(* IEC 61131-3 sources: daoli-st-library/DL_Process (part 56) *)

(* ---- FB_DL_TireCureBlowdownWatch.st ---- *)
(*
  Name: FB_DL_TireCureBlowdownWatch
  Category: DL_Process
  Version: 1.0.0
  Round: R91 / 2026-11-25
  开源溯源：clean-room 自研（族 轮胎硫化，ST 开源生态实测 0 命中，无外部代码引入）
  功能：1) 按固定观察窗累计两个量：冷凝水总量 _fAccumKg 与排凝阀动作次数 _iAccumAct，
           窗口到点后按「单位动作排水量」比对：
           ratio = 累计冷凝水 / (动作次数 × 单次期望排水量)。
        2) 双向故障判别：
           ① 比值过高（> fBlockRatio）或窗口内动作次数为零而冷凝水已超限 → 判排凝阀堵塞（码 0322 / 0324），
              即水积在腔内排不出去，会稀释硫化温度场并造成胶囊局部过冷；
           ② 比值过低（< fLeakRatio）→ 判排凝阀泄漏（码 0323），即阀频繁动作但排水极少，
              说明阀芯未关严、蒸汽直排，属能耗与安全问题。
        3) 窗口自复位由 TON 的 IN := xEnable AND NOT tonWin.Q 驱动（R188），
           窗口到点仅置 Q 一拍，用于「判定 + 清累计」的一次性动作，不靠外部沿清零。
  边界条件：1) 非有限值闸：冷凝水量、期望排水量、两个比值阈值、窗口先过
           NOT(x > -DL_BIG AND x < DL_BIG)，同时拦 NaN 与 Inf；命中即锁码 0326 进故障相，
           绝不把 NaN 累加进窗口（NaN 一旦进入累计器，整个窗口乃至后续窗口永久污染，R19）。
        2) 分母零闸：比值式分母 = 动作次数 × 单次期望排水量，动作次数为零时走独立判据（码 0324），
           单次期望排水量 fExpectKgPerAct 必须 > DL_EPS 否则锁码 0325（判据全体失效）。
        3) 阈值域闸：须满足 0.0 < fLeakRatio < fBlockRatio，否则两向判据重叠、必有一向永不触发，
           越域锁码 0325。
        4) 累计器安全：非有限值命中时把两个累计器一并清零（码 0326 已锁存），
           并中止本窗口的判定，防污染值跨窗口传播。
        5) 定时器周期刷新（R7）：窗口 TON 与两个边沿实例全部在 CASE 之外无条件调用。
        6) 故障解除路径：故障相内 xReset 上升沿 AND NOT xFault AND 入参/组态合法 → 清锁存回正常，
           回正常后窗口与累计器全部重新起算（不自恢复）。
        7) 状态机兜底：CASE 全态覆盖 + ELSE 强制回故障相并置码 0328、清全部输出。
        8) 输出安全初值（R25）：xBlocked / xLeaking 初值 FALSE，fRatioPct 初值 0.0，正常相显式赋值。
  量纲自证：ratio = (kg) / (无因次 * kg) = 无因次 [-]；fRatioPct = 无因次 * 100 = 百分数 [%]；
           fAccumKg 为累计质量 [kg]，nAccumAct 为动作次数（计数，无量纲）[count]。
  码表 Error codes（本件子带 0091_032x，故障级一律 3 行内置 _uFault/_bFault/_eState）:
    16#0091_0321 信息级：观察窗累计中，尚未判定（不置故障位）
    16#0091_0322 故障级：排凝阀堵塞（单位动作排水量比值过高）
    16#0091_0323 故障级：排凝阀泄漏（单位动作排水量比值过低，蒸汽直排）
    16#0091_0324 故障级：窗口内动作次数为零但冷凝水超限（阀未动作）
    16#0091_0325 故障级：组态越域（期望排水量/比值阈值/窗口非法）
    16#0091_0326 故障级：入参非有限（NaN 或 Inf），累计器已清
    16#0091_0327 故障级：外部故障输入 xFault
    16#0091_0328 故障级：状态机落 ELSE 兜底（非法相位 ID）

  修订历史 Revision :
    2026-11-25  v1.0.0  R91 首版
*)

TYPE E_DL_TcsBlowdownState :
(
    eTcsBdNormal  := 0,     // 正常：窗口比值在带内 / Normal, window ratio within the band
    eTcsBdBlocked := 10,    // 排凝阀堵塞：水排不出去 / Blocked blowdown valve, water cannot be discharged
    eTcsBdLeaking := 20,    // 排凝阀泄漏：蒸汽直排 / Leaking blowdown valve, steam blows through
    eTcsBdFault   := 90     // 故障：入参/组态非法，锁存待解除 / Fault, invalid input, latched
);
END_TYPE

FUNCTION_BLOCK FB_DL_TireCureBlowdownWatch
VAR_INPUT
    xEnable         : BOOL;   // 监视使能 [bool] / Monitoring enable [bool]
    xReset          : BOOL;   // 故障复位（上升沿有效）[bool] / Fault reset, rising edge [bool]
    xFault          : BOOL;   // 外部故障汇总 [bool] / External fault aggregate [bool]
    xCyclePulse     : BOOL;   // 周期完成脉冲（每个模压周期一个脉冲）[bool] / Cycle-complete pulse [bool]
    fCondensateKg   : REAL;   // 本周期冷凝水量增量 [kg] / Condensate increment of this cycle [kg]
    nActCount       : INT;    // 本周期排凝阀动作次数 [count] / Blowdown valve actuations this cycle [count]
    fExpectKgPerAct : REAL;   // 单次动作期望排水量 [kg/act] / Expected discharge per actuation [kg/act]
    fBlockRatio     : REAL;   // 堵塞判定比值上限 [-] / Blockage upper ratio limit [-]
    fLeakRatio      : REAL;   // 泄漏判定比值下限 [-] / Leakage lower ratio limit [-]
    tWindow         : TIME;   // 观察窗时长 [TIME] / Observation window duration [TIME]
END_VAR
VAR_OUTPUT
    fRatioPct       : REAL;   // 窗口单位动作排水量比值（百分数显示）[%] / Window ratio, percent display [%]
    fAccumKg        : REAL;   // 窗口累计冷凝水量 [kg] / Accumulated condensate in the window [kg]
    nAccumAct       : INT;    // 窗口累计动作次数 [count] / Accumulated actuations in the window [count]
    xBlocked        : BOOL;   // 堵塞标志 [bool] / Blockage flag [bool]
    xLeaking        : BOOL;   // 泄漏标志 [bool] / Leakage flag [bool]
    xWindowDone     : BOOL;   // 窗口到点脉冲（单拍）[bool] / Window-complete single-shot flag [bool]
    eState          : E_DL_TcsBlowdownState;   // 状态出口，段尾单点映射 / State outlet, single-point mapped
    nErrId          : UDINT;  // 事件码，0 = 无事件 / Event code, 0 = none
END_VAR
VAR
    tonWin          : TON;    // 观察窗定时（自复位由 IN 取反驱动，R188）[TIME] / Observation window timer
    rtCycle         : R_TRIG; // 周期脉冲上升沿检测 [bool] / Cycle pulse rising edge detector
    rtReset         : R_TRIG; // 复位上升沿检测 [bool] / Reset rising edge detector
    _eState         : E_DL_TcsBlowdownState := E_DL_TcsBlowdownState.eTcsBdNormal;   // 内部相位（CASE 唯一写入目标）
    _fAccumKg       : REAL := 0.0;   // 窗口累计冷凝水量 [kg] / Accumulated condensate [kg]
    _iAccumAct      : INT := 0;      // 窗口累计动作次数 [count] / Accumulated actuations [count]
    _fRatioRaw      : REAL := 0.0;   // 窗口比值原始值（无因次）[-] / Raw window ratio [-]
    _fRatioRawPct   : REAL := 0.0;   // 窗口比值百分数原始值 [%] / Raw window ratio in percent [%]
    _bFinOk         : BOOL := FALSE; // 实值入参有限性总闸结果 / Finiteness gate aggregate result
    _bCfgOk         : BOOL := FALSE; // 阈值与窗口组态域闸结果 / Threshold and window domain gate result
    _bJudgeThis     : BOOL := FALSE; // 本拍需执行窗口判定（窗口到点）[bool] / Judge this cycle flag
    _bBlockedL      : BOOL := FALSE; // 堵塞锁存位 [bool] / Latched blockage flag
    _bLeakingL      : BOOL := FALSE; // 泄漏锁存位 [bool] / Latched leakage flag
    _bFault         : BOOL := FALSE; // 故障锁存位 [bool] / Latched fault flag
    _uInfo          : UDINT := 16#0000_0000;   // 信息码，每拍重算 / Info code, recomputed every cycle
    _uFault         : UDINT := 16#0000_0000;   // 故障码锁存 / Latched fault code
END_VAR
VAR CONSTANT
    DL_EPS         : REAL := 1.0E-9;      // 数值零闸阈值 [-] / Numeric zero gate threshold [-]
    DL_BIG         : REAL := 1.0E12;      // 非有限值闸量级上限 [-] / Finiteness gate magnitude [-]
    DL_PCT         : REAL := 100.0;       // 百分比换算因子 [%] / Percent conversion factor [%]
    DL_RATIO_HI    : REAL := 1000.0;      // 比值显示上限 [-] / Ratio display ceiling [-]
    DL_ACCUM_HI_KG : REAL := 10000.0;     // 累计水量物理上限 [kg] / Accumulated mass upper bound [kg]
    DL_ACT_HI      : INT := 100000;       // 累计次数物理上限 [count] / Accumulation count upper bound [count]
    DL_WATER_MIN_KG : REAL := 0.001;      // 判定「有冷凝水」的最小累计量 [kg] / Minimum condensate to judge [kg]
END_VAR

(* —— 段 0：单拍量预清零（锁存量 _uFault/_bFault/_bBlockedL/_bLeakingL/_fAccumKg/_iAccumAct 不入清单，R187①） —— *)
(*     注：_fRatioRaw / _fRatioRawPct 为「上一窗口判定值」保持量，故意不在此清零，供面板持续显示。 *)
_uInfo := 16#0000_0000;                     // 信息码每拍重算 / Info code recomputed
nErrId := 16#0000_0000;                     // 事件码缺省无事件 / Event code defaults to none

(* —— 段 1：非有限值闸与组态域闸（R19：不把 NaN 累加进窗口） —— *)
_bFinOk := (fCondensateKg > -DL_BIG) AND (fCondensateKg < DL_BIG)
           AND (fExpectKgPerAct > -DL_BIG) AND (fExpectKgPerAct < DL_BIG)
           AND (fBlockRatio > -DL_BIG) AND (fBlockRatio < DL_BIG)
           AND (fLeakRatio > -DL_BIG) AND (fLeakRatio < DL_BIG);
_bCfgOk := (fExpectKgPerAct > DL_EPS)                     // 期望单次排水量必须为正（比值分母）
           AND (fLeakRatio > DL_EPS)                       // 泄漏下限必须为正
           AND (fBlockRatio > fLeakRatio)                   // 堵塞上限必须严格大于泄漏下限
           AND (fBlockRatio <= DL_RATIO_HI)                // 上限须在显示域内
           AND (nActCount >= 0)                            // 动作次数不得为负
           AND (tWindow > T#0S);                           // 观察窗必须为正

(* —— 段 2：边沿与窗口定时器无条件周期刷新（R7：调用语句不得置于 IF/CASE 内） —— *)
rtCycle(CLK := xCyclePulse);                                                    // 周期脉冲上升沿，每拍必调
rtReset(CLK := xReset);                                                         // 复位上升沿，每拍必调
tonWin(IN := xEnable AND (NOT tonWin.Q), PT := tWindow);                        // 观察窗自复位（R188）
_bJudgeThis := tonWin.Q;                                                        // 窗口到点：本拍执行判定

(* —— 段 3：窗口累计（仅在有限值且组态合法时累加，防污染跨窗口传播） —— *)
IF rtCycle.Q AND _bFinOk AND _bCfgOk THEN
    _fAccumKg := _fAccumKg + fCondensateKg;             // 累计冷凝水 [kg]
    _iAccumAct := _iAccumAct + nActCount;               // 累计动作次数 [count]
END_IF

(* —— 段 4：全局故障拦截（优先级最高；已锁存则不再改写码值，禁同拍抹除） —— *)
IF xFault AND (NOT _bFault) THEN
    _uFault := 16#0091_0327;                // 故障级：外部故障输入
    _bFault := TRUE;                        // 锁存（3 行内置，R45 配对）
    _eState := E_DL_TcsBlowdownState.eTcsBdFault;
END_IF
IF (NOT _bFinOk) AND (NOT _bFault) THEN
    _uFault := 16#0091_0326;                // 故障级：入参非有限
    _bFault := TRUE;                        // 锁存
    _fAccumKg := 0.0;                       // 累计器清（防污染跨窗口）
    _iAccumAct := 0;                        // 计数清
    _eState := E_DL_TcsBlowdownState.eTcsBdFault;
END_IF
IF (NOT _bCfgOk) AND _bFinOk AND (NOT _bFault) THEN
    _uFault := 16#0091_0325;                // 故障级：组态越域（独立成因，R190）
    _bFault := TRUE;                        // 锁存
    _eState := E_DL_TcsBlowdownState.eTcsBdFault;
END_IF

(* —— 段 5：相位机（只做迁移与锁存；出口在段 7 单点映射） —— *)
CASE _eState OF

E_DL_TcsBlowdownState.eTcsBdNormal:
    IF NOT xEnable THEN
        _uInfo := 16#0091_0321;             // 信息级：监视关闭，累计冻结（不置故障位）
    ELSIF _bJudgeThis THEN
        IF (_iAccumAct <= 0) AND (_fAccumKg > DL_WATER_MIN_KG) THEN
            _uFault := 16#0091_0324;        // 故障级：动作次数为零但水已积（阀未动作）
            _bBlockedL := TRUE;             // 堵塞锁存
            _eState := E_DL_TcsBlowdownState.eTcsBdBlocked;
        ELSIF (_iAccumAct > 0) AND (ABS(fExpectKgPerAct * INT_TO_REAL(_iAccumAct)) > DL_EPS) THEN
            _fRatioRaw := _fAccumKg / (fExpectKgPerAct * INT_TO_REAL(_iAccumAct));   // 比值 [-]
            _fRatioRawPct := _fRatioRaw * DL_PCT;                                    // 百分数显示 [%]
            IF _fRatioRaw > fBlockRatio THEN
                _uFault := 16#0091_0322;    // 故障级：比值过高，阀堵塞
                _bBlockedL := TRUE;         // 堵塞锁存
                _eState := E_DL_TcsBlowdownState.eTcsBdBlocked;
            ELSIF _fRatioRaw < fLeakRatio THEN
                _uFault := 16#0091_0323;    // 故障级：比值过低，阀泄漏
                _bLeakingL := TRUE;         // 泄漏锁存
                _eState := E_DL_TcsBlowdownState.eTcsBdLeaking;
            ELSE
                _uInfo := 16#0091_0321;     // 信息级：窗口比值合格，进入下一窗口
            END_IF
        ELSE
            _uInfo := 16#0091_0321;         // 信息级：窗口内无有效动作，无法判定
        END_IF
        _fAccumKg := 0.0;                   // 窗口结束：累计清零（判定后统一清，R187 同拍不抹判定）
        _iAccumAct := 0;                    // 窗口结束：计数清零
    ELSE
        _uInfo := 16#0091_0321;             // 信息级：累计中，尚未判定
    END_IF

E_DL_TcsBlowdownState.eTcsBdBlocked:
    IF rtReset.Q THEN
        _bBlockedL := FALSE;                // 解除路径：复位上升沿（可达，R188）
        _uFault := 16#0000_0000;            // 清锁存码
        _fAccumKg := 0.0;                   // 累计器重新起算
        _iAccumAct := 0;                    // 计数重新起算
        _eState := E_DL_TcsBlowdownState.eTcsBdNormal;
    END_IF

E_DL_TcsBlowdownState.eTcsBdLeaking:
    IF rtReset.Q THEN
        _bLeakingL := FALSE;                // 解除路径：复位上升沿（可达，R188）
        _uFault := 16#0000_0000;            // 清锁存码
        _fAccumKg := 0.0;                   // 累计器重新起算
        _iAccumAct := 0;                    // 计数重新起算
        _eState := E_DL_TcsBlowdownState.eTcsBdNormal;
    END_IF

E_DL_TcsBlowdownState.eTcsBdFault:
    IF rtReset.Q AND (NOT xFault) AND _bFinOk AND _bCfgOk THEN
        _bFault := FALSE;                   // 解除路径：复位沿 + 外部故障消失 + 入参/组态合法（可达，R188）
        _uFault := 16#0000_0000;            // 清锁存码
        _fAccumKg := 0.0;                   // 累计器重新起算
        _iAccumAct := 0;                    // 计数重新起算
        _eState := E_DL_TcsBlowdownState.eTcsBdNormal;
    END_IF

ELSE
    _uFault := 16#0091_0328;                // 故障级：非法相位 ID 兜底
    _bFault := TRUE;                        // 锁存
    _bBlockedL := FALSE;                    // 各级锁存清
    _bLeakingL := FALSE;
    _fAccumKg := 0.0;                       // 累计器清
    _iAccumAct := 0;
    _eState := E_DL_TcsBlowdownState.eTcsBdFault;             // 强制回故障相

END_CASE

(* —— 段 6：后置段（累计器域兜底：非有限或越量级即清零，防污染跨窗口） —— *)
IF NOT (_fAccumKg > -DL_BIG AND _fAccumKg < DL_BIG) THEN
    _fAccumKg := 0.0;                       // 内部状态自检：非有限即清零
END_IF
IF _fAccumKg > DL_ACCUM_HI_KG THEN
    _fAccumKg := DL_ACCUM_HI_KG;            // 越物理上限钳制，防累计器发散
END_IF
IF _iAccumAct > DL_ACT_HI THEN
    _iAccumAct := DL_ACT_HI;                // 越计数上限钳制，防整型溢出
END_IF
IF _iAccumAct < 0 THEN
    _iAccumAct := 0;                        // 负计数属异常，归零（不参与比值分母）
END_IF

(* —— 段 7：出口单点映射（名实同源；锁存位一律由状态导出，故障侧全清） —— *)
fRatioPct := LIMIT(0.0, _fRatioRawPct, DL_RATIO_HI * DL_PCT);                     // 比值百分数钳显示域 [%]
fAccumKg := MIN(_fAccumKg, DL_ACCUM_HI_KG);                                       // 累计量出口（已钳，单点写）
nAccumAct := _iAccumAct;                                                          // 累计次数出口
xBlocked := _bBlockedL AND (NOT _bFault);                                         // 堵塞位出口
xLeaking := _bLeakingL AND (NOT _bFault);                                         // 泄漏位出口
xWindowDone := _bJudgeThis;                                                       // 窗口到点单拍脉冲出口
eState := _eState;                                                                // 状态出口单点映射
IF _bFault OR _bBlockedL OR _bLeakingL THEN
    nErrId := _uFault;                      // 故障码锁存回放（不在故障相按当下输入重推断）
ELSE
    nErrId := _uInfo;                       // 信息码
END_IF

END_FUNCTION_BLOCK

(* ---- FB_DL_TireCureMoldTempWatch.st ---- *)
(*
  Name: FB_DL_TireCureMoldTempWatch
  Category: DL_Process
  Version: 1.0.0
  Round: R91 / 2026-11-25
  开源溯源：clean-room 自研（族 轮胎硫化，ST 开源生态实测 0 命中，无外部代码引入）
  功能：1) 上下模温差监视：dT = |上模温 − 下模温|，两级判据并行且各自去抖：
           超过 fDeltaWarnK 进预警（信息级码 0312），超过 fDeltaMaxK 进报警（故障级码 0314）。
           上下模温差过大意味着单侧加热回路能力不足，会造成硫化程度沿胎圈-胎面方向不均。
        2) 加热失效判据：由实测上模温按周期折算温升速率 r = dT/dt [K/min]，
           r 的绝对值低于 fHeatRateMinKmin 且持续一个去抖窗，判加热失效（码 0315）——
           这是热电偶脱落与固态继电器击穿共有的实测特征（温度「不动」）。
        3) 趋势方向输出 nTrend：+1 上升、0 平稳、-1 下降，由本拍与上拍上模温差按
           DL_TREND_K 死区判定，供上层画趋势箭头与判断「是否正在爬温」。
  边界条件：1) 非有限值闸：温度、阈值、周期先过 NOT(x > -DL_BIG AND x < DL_BIG)，同时拦 NaN 与 Inf；
           命中即锁码 0317 进故障相 —— 绝不让 NaN 参与温差与速率计算
           （NaN 比较恒假会把「测点断线」伪装成「温差正常、速率正常」，R19）。
        2) 周期入参闸（R21）：fCycleS <= 0.0 或非有限时改用缺省 DL_CYCLE_DEF = 0.1 s，
           温升速率的折算依赖该值，故必须显式声明（码 0317 同码归因，内部成员分离）。
        3) 阈值域闸：须满足 0.0 < fDeltaWarnK < fDeltaMaxK 且 fHeatRateMinKmin > DL_EPS，
           越域锁码 0317（预警/报警两级重叠或倒置会让某级永不触发）。
        4) 快照闸：首拍 _bPrevValid = FALSE 时不判速率与趋势，避免上电「上拍温度 = 0」
           造成的假加热失效。
        5) 定时器周期刷新（R7）：三个 TON 与复位边沿全部在 CASE 之外无条件调用。
        6) 故障解除路径：故障相内 xReset 上升沿 AND NOT xFault AND 入参/组态合法 → 清锁存回正常，
           回正常需重新积累去抖窗（不自恢复）。
        7) 状态机兜底：CASE 全态覆盖 + ELSE 强制回故障相并置码 0318、清全部输出。
        8) 输出安全初值（R25）：xWarn / xAlarm / xHeatFail 初值 FALSE，nTrend 初值 0，
           正常相显式赋值。
  量纲自证：dT = |(degC) − (degC)| = (K)；趋势死区 DL_TREND_K 为 [K]，与温差同量纲；
           r = dT[K] / fCycleS[s] * 60[s/min] = K/min，与 fHeatRateMinKmin 同量纲。
  码表 Error codes（本件子带 0091_031x，故障级一律 3 行内置 _uFault/_bFault/_eState）:
    16#0091_0311 信息级：使能关闭，监视冻结（不置故障位）
    16#0091_0312 信息级：上下模温差已超预警阈值，尚在去抖窗内（不置故障位）
    16#0091_0313 故障级：上下模温差超预警阈值（去抖确认）
    16#0091_0314 故障级：上下模温差超上限阈值（去抖确认）
    16#0091_0315 故障级：加热失效（温升速率绝对值低于下限）
    16#0091_0316 故障级：外部故障输入 xFault
    16#0091_0317 故障级：入参非有限或阈值/周期组态越域
    16#0091_0318 故障级：状态机落 ELSE 兜底（非法相位 ID）

  修订历史 Revision :
    2026-11-25  v1.0.0  R91 首版
*)

TYPE E_DL_TcsMoldTempState :
(
    eTcsMoldNormal   := 0,    // 正常：温差与速率均在带内 / Normal, difference and rate within limits
    eTcsMoldWarn     := 10,   // 预警：温差超预警阈值（已去抖）/ Warning, difference over the warning limit
    eTcsMoldAlarm    := 20,   // 报警：温差超上限阈值（已去抖）/ Alarm, difference over the upper limit
    eTcsMoldHeatFail := 30,   // 加热失效：温升速率不足（已去抖）/ Heat failure, rate below the limit
    eTcsMoldFault    := 90    // 故障：入参/组态非法，锁存待解除 / Fault, invalid input, latched
);
END_TYPE

FUNCTION_BLOCK FB_DL_TireCureMoldTempWatch
VAR_INPUT
    xEnable        : BOOL;    // 监视使能 [bool] / Monitoring enable [bool]
    xReset         : BOOL;    // 故障复位（上升沿有效）[bool] / Fault reset, rising edge [bool]
    xFault         : BOOL;    // 外部故障汇总 [bool] / External fault aggregate [bool]
    fUpperMoldC    : REAL;    // 上模温度 [degC] / Upper mold temperature [degC]
    fLowerMoldC    : REAL;    // 下模温度 [degC] / Lower mold temperature [degC]
    fDeltaWarnK    : REAL;    // 温差预警阈值 [K] / Temperature difference warning threshold [K]
    fDeltaMaxK     : REAL;    // 温差上限阈值 [K] / Temperature difference upper limit [K]
    fHeatRateMinKmin : REAL;  // 允许最小温升速率（绝对值）[K/min] / Minimum absolute heating rate [K/min]
    fCycleS        : REAL;    // 任务周期 [s] / Task cycle time [s]
    tDebounce      : TIME;    // 判据去抖窗 [TIME] / Criteria debounce window [TIME]
END_VAR
VAR_OUTPUT
    fDeltaK        : REAL;    // 上下模温差绝对值 [K] / Absolute mold temperature difference [K]
    fRateKmin      : REAL;    // 上模温升速率（带符号）[K/min] / Upper mold heating rate, signed [K/min]
    nTrend         : INT;     // 趋势方向 +1 升 / 0 平 / -1 降 [dir] / Trend direction +1/0/-1 [dir]
    xWarn          : BOOL;    // 预警位（信息级）[bool] / Warning flag, information grade [bool]
    xAlarm         : BOOL;    // 报警位（故障级）[bool] / Alarm flag, fault grade [bool]
    xHeatFail      : BOOL;    // 加热失效位 [bool] / Heat failure flag [bool]
    eState         : E_DL_TcsMoldTempState;   // 状态出口，段尾单点映射 / State outlet, single-point mapped
    nErrId         : UDINT;   // 事件码，0 = 无事件 / Event code, 0 = none
END_VAR
VAR
    tonWarn        : TON;     // 温差预警去抖定时 [TIME] / Difference warning debounce timer
    tonAlarm       : TON;     // 温差报警去抖定时 [TIME] / Difference alarm debounce timer
    tonHeat        : TON;     // 加热失效去抖定时 [TIME] / Heat failure debounce timer
    rtReset        : R_TRIG;  // 复位上升沿检测 [bool] / Reset rising edge detector
    _eState        : E_DL_TcsMoldTempState := E_DL_TcsMoldTempState.eTcsMoldNormal;   // 内部相位（CASE 唯一写入目标）
    _fUpperPrevC   : REAL := 0.0;   // 上拍上模温度快照 [degC] / Previous-cycle upper mold temperature [degC]
    _bPrevValid    : BOOL := FALSE; // 温度快照有效位（首拍为假）/ Temperature snapshot validity, false on first cycle
    _fCycleUseS    : REAL := 0.1;   // 实际使用的周期值 [s] / Cycle time actually used [s]
    _fDeltaRawK    : REAL := 0.0;   // 温差原始值 [K] / Raw temperature difference [K]
    _fRateRawKmin  : REAL := 0.0;   // 温升速率原始值 [K/min] / Raw heating rate [K/min]
    _bFinOk        : BOOL := FALSE; // 实值入参有限性总闸结果 / Finiteness gate aggregate result
    _bCfgOk        : BOOL := FALSE; // 阈值与周期组态域闸结果 / Threshold and cycle domain gate result
    _bWarnRaw      : BOOL := FALSE; // 温差预警原始判据 [bool] / Raw difference warning criterion
    _bAlarmRaw     : BOOL := FALSE; // 温差报警原始判据 [bool] / Raw difference alarm criterion
    _bHeatRaw      : BOOL := FALSE; // 加热失效原始判据 [bool] / Raw heat failure criterion
    _bWarnL        : BOOL := FALSE; // 预警锁存位 [bool] / Latched warning flag
    _bAlarmL       : BOOL := FALSE; // 报警锁存位 [bool] / Latched alarm flag
    _bHeatL        : BOOL := FALSE; // 加热失效锁存位 [bool] / Latched heat-failure flag
    _bFault        : BOOL := FALSE; // 故障锁存位 [bool] / Latched fault flag
    _uInfo         : UDINT := 16#0000_0000;   // 信息码，每拍重算 / Info code, recomputed every cycle
    _uFault        : UDINT := 16#0000_0000;   // 故障码锁存 / Latched fault code
END_VAR
VAR CONSTANT
    DL_EPS         : REAL := 1.0E-9;      // 数值零闸阈值 [-] / Numeric zero gate threshold [-]
    DL_BIG         : REAL := 1.0E12;      // 非有限值闸量级上限 [-] / Finiteness gate magnitude [-]
    DL_CYCLE_DEF   : REAL := 0.1;         // 缺省任务周期 [s] / Default task cycle time [s]
    DL_CYCLE_MIN   : REAL := 0.001;       // 周期合理下限 [s] / Cycle time reasonable low bound [s]
    DL_CYCLE_MAX   : REAL := 10.0;        // 周期合理上限 [s] / Cycle time reasonable high bound [s]
    DL_SEC_PER_MIN : REAL := 60.0;        // 分钟到秒的时基折算 [s/min] / Seconds per minute [s/min]
    DL_TREND_K     : REAL := 0.2;         // 趋势判定死区 [K] / Trend dead band [K]
    DL_DELTA_HI    : REAL := 500.0;       // 温差物理上限 [K] / Temperature difference upper bound [K]
    DL_RATE_HI     : REAL := 100.0;       // 温升速率物理上限 [K/min] / Heating rate upper bound [K/min]
    DL_T_SPAN      : REAL := 500.0;       // 温度量级闸跨度 [degC] / Temperature magnitude gate span [degC]
END_VAR

(* —— 段 0：单拍量预清零（锁存量 _uFault/_bFault/_bWarnL/_bAlarmL/_bHeatL 不入清单，R187①） —— *)
_uInfo := 16#0000_0000;                     // 信息码每拍重算 / Info code recomputed
nErrId := 16#0000_0000;                     // 事件码缺省无事件 / Event code defaults to none

(* —— 段 1：周期入参闸（R21）与非有限值闸（R19） —— *)
_bFinOk := (fUpperMoldC > -DL_BIG) AND (fUpperMoldC < DL_BIG)
           AND (fLowerMoldC > -DL_BIG) AND (fLowerMoldC < DL_BIG)
           AND (fDeltaWarnK > -DL_BIG) AND (fDeltaWarnK < DL_BIG)
           AND (fDeltaMaxK > -DL_BIG) AND (fDeltaMaxK < DL_BIG)
           AND (fHeatRateMinKmin > -DL_BIG) AND (fHeatRateMinKmin < DL_BIG)
           AND (fCycleS > -DL_BIG) AND (fCycleS < DL_BIG);
_bCfgOk := (fDeltaWarnK > DL_EPS)                       // 预警阈值必须为正
           AND (fDeltaMaxK > fDeltaWarnK)               // 上限必须严格大于预警
           AND (fDeltaMaxK <= DL_DELTA_HI)              // 上限须在物理域内
           AND (fHeatRateMinKmin > DL_EPS)              // 速率下限必须为正
           AND (ABS(fUpperMoldC) <= DL_T_SPAN)          // 温度量级闸
           AND (ABS(fLowerMoldC) <= DL_T_SPAN)
           AND (fCycleS >= DL_CYCLE_MIN) AND (fCycleS <= DL_CYCLE_MAX)
           AND (tDebounce > T#0S);                      // 去抖窗必须为正

IF _bCfgOk THEN
    _fCycleUseS := fCycleS;                 // 合法周期原值使用
ELSE
    _fCycleUseS := DL_CYCLE_DEF;            // 非法周期一律用缺省 0.1 s（组态闸在段 5 统一判）
END_IF

(* —— 段 2：判据派生（原始值；快照闸保证首拍不判速率） —— *)
_fDeltaRawK := ABS(fUpperMoldC - fLowerMoldC);                                    // 上下模温差 [K]
IF _bPrevValid AND _bFinOk THEN
    _fRateRawKmin := (fUpperMoldC - _fUpperPrevC) / _fCycleUseS * DL_SEC_PER_MIN; // 温升速率 [K/min]
ELSE
    _fRateRawKmin := 0.0;                   // 首拍无快照：速率置零（不据此判失效）
END_IF
_bWarnRaw := _bFinOk AND _bCfgOk AND xEnable AND (_fDeltaRawK > fDeltaWarnK);
_bAlarmRaw := _bFinOk AND _bCfgOk AND xEnable AND (_fDeltaRawK > fDeltaMaxK);
_bHeatRaw := _bFinOk AND _bCfgOk AND xEnable AND _bPrevValid
             AND (ABS(_fRateRawKmin) < fHeatRateMinKmin);

(* —— 段 3：定时器与边沿无条件周期刷新（R7：调用语句不得置于 IF/CASE 内） —— *)
rtReset(CLK := xReset);                                                     // 复位上升沿，每拍必调
tonWarn(IN := _bWarnRaw AND (NOT _bFault), PT := tDebounce);                 // 温差预警去抖
tonAlarm(IN := _bAlarmRaw AND (NOT _bFault), PT := tDebounce);               // 温差报警去抖
tonHeat(IN := _bHeatRaw AND (NOT _bFault), PT := tDebounce);                 // 加热失效去抖

(* —— 段 4：全局故障拦截（优先级最高；已锁存则不再改写码值，禁同拍抹除） —— *)
IF xFault AND (NOT _bFault) THEN
    _uFault := 16#0091_0316;                // 故障级：外部故障输入
    _bFault := TRUE;                        // 锁存（3 行内置，R45 配对）
    _eState := E_DL_TcsMoldTempState.eTcsMoldFault;
END_IF
IF ((NOT _bFinOk) OR (NOT _bCfgOk)) AND (NOT _bFault) THEN
    _uFault := 16#0091_0317;                // 故障级：入参非有限或组态越域（内部成员已分离）
    _bFault := TRUE;                        // 锁存
    _eState := E_DL_TcsMoldTempState.eTcsMoldFault;
END_IF

(* —— 段 5：相位机（只做迁移与锁存；出口在段 7 单点映射） —— *)
CASE _eState OF

E_DL_TcsMoldTempState.eTcsMoldNormal:
    IF NOT xEnable THEN
        _uInfo := 16#0091_0311;             // 信息级：使能关闭，监视冻结（不置故障位）
    ELSIF tonAlarm.Q THEN
        _uFault := 16#0091_0314;            // 故障级：温差超上限（去抖确认）
        _bAlarmL := TRUE;                   // 报警锁存
        _eState := E_DL_TcsMoldTempState.eTcsMoldAlarm;
    ELSIF tonHeat.Q THEN
        _uFault := 16#0091_0315;            // 故障级：加热失效（去抖确认）
        _bHeatL := TRUE;                    // 加热失效锁存
        _eState := E_DL_TcsMoldTempState.eTcsMoldHeatFail;
    ELSIF tonWarn.Q THEN
        _uFault := 16#0091_0313;            // 故障级：温差超预警（去抖确认）
        _bWarnL := TRUE;                    // 预警锁存
        _eState := E_DL_TcsMoldTempState.eTcsMoldWarn;
    ELSIF _bWarnRaw THEN
        _uInfo := 16#0091_0312;             // 信息级：超预警阈值但尚在去抖窗内
    END_IF

E_DL_TcsMoldTempState.eTcsMoldWarn:
    IF NOT xEnable THEN
        _uInfo := 16#0091_0311;             // 信息级：使能关闭，监视冻结
        _bWarnL := FALSE;                   // 失能即清预警锁存
        _eState := E_DL_TcsMoldTempState.eTcsMoldNormal;
    ELSIF tonAlarm.Q THEN
        _uFault := 16#0091_0314;            // 故障级：温差升级到上限
        _bAlarmL := TRUE;                   // 报警锁存
        _eState := E_DL_TcsMoldTempState.eTcsMoldAlarm;
    ELSIF NOT _bWarnRaw THEN
        _bWarnL := FALSE;                   // 判据自行消失：清预警锁存回正常（无需复位）
        _eState := E_DL_TcsMoldTempState.eTcsMoldNormal;
    END_IF

E_DL_TcsMoldTempState.eTcsMoldAlarm:
    IF rtReset.Q THEN
        _bAlarmL := FALSE;                  // 解除路径：复位上升沿（可达，R188）
        _uFault := 16#0000_0000;            // 清锁存码
        _eState := E_DL_TcsMoldTempState.eTcsMoldNormal;
    END_IF

E_DL_TcsMoldTempState.eTcsMoldHeatFail:
    IF rtReset.Q THEN
        _bHeatL := FALSE;                   // 解除路径：复位上升沿（可达，R188）
        _uFault := 16#0000_0000;            // 清锁存码
        _bPrevValid := FALSE;               // 强制重新取快照，避免旧快照立刻再判失效
        _eState := E_DL_TcsMoldTempState.eTcsMoldNormal;
    END_IF

E_DL_TcsMoldTempState.eTcsMoldFault:
    IF rtReset.Q AND (NOT xFault) AND _bFinOk AND _bCfgOk THEN
        _bFault := FALSE;                   // 解除路径：复位沿 + 外部故障消失 + 入参/组态合法（可达，R188）
        _uFault := 16#0000_0000;            // 清锁存码
        _bPrevValid := FALSE;               // 强制重新取快照
        _eState := E_DL_TcsMoldTempState.eTcsMoldNormal;
    END_IF

ELSE
    _uFault := 16#0091_0318;                // 故障级：非法相位 ID 兜底
    _bFault := TRUE;                        // 锁存
    _bWarnL := FALSE;                       // 各级锁存清
    _bAlarmL := FALSE;
    _bHeatL := FALSE;
    _eState := E_DL_TcsMoldTempState.eTcsMoldFault;           // 强制回故障相

END_CASE

(* —— 段 6：后置段（温度快照在迁移判断之后统一更新，禁在分支内散写） —— *)
IF _bFinOk THEN
    _fUpperPrevC := fUpperMoldC;            // 快照更新（仅有限值可信时才更新）
    _bPrevValid := TRUE;                    // 快照自此有效
ELSE
    _bPrevValid := FALSE;                   // 非有限值使快照失效，防污染下一拍速率判据
END_IF

(* —— 段 7：出口单点映射（名实同源；锁存位一律由状态导出，故障侧全清） —— *)
fDeltaK := LIMIT(0.0, _fDeltaRawK, DL_DELTA_HI);                                  // 温差出口钳物理域 [K]
fRateKmin := LIMIT(-DL_RATE_HI, _fRateRawKmin, DL_RATE_HI);                       // 速率出口钳物理域 [K/min]
IF _fRateRawKmin > DL_TREND_K THEN
    nTrend := 1;                            // 上升
ELSIF _fRateRawKmin < -DL_TREND_K THEN
    nTrend := -1;                           // 下降
ELSE
    nTrend := 0;                            // 平稳（死区内）
END_IF
xWarn := _bWarnL AND (NOT _bFault);                                        // 预警位出口
xAlarm := _bAlarmL AND (NOT _bFault);                                      // 报警位出口
xHeatFail := _bHeatL AND (NOT _bFault);                                    // 加热失效出口
eState := _eState;                                                         // 状态出口单点映射
IF _bFault OR _bAlarmL OR _bHeatL OR _bWarnL THEN
    nErrId := _uFault;                      // 故障码锁存回放（不在故障相按当下输入重推断）
ELSE
    nErrId := _uInfo;                       // 信息码
END_IF

END_FUNCTION_BLOCK

(* ---- FB_DL_TireCurePressSeq.st ---- *)
(*
  Name: FB_DL_TireCurePressSeq
  Category: DL_Process
  Version: 1.0.0
  Round: R91 / 2026-11-25
  开源溯源：clean-room 自研（族 轮胎硫化，ST 开源生态实测 0 命中，无外部代码引入）
  功能：1) 硫化机合模序状态机，十相推进（含故障相）：
           待机 → 装胎 → 合模 → 一次定型 → 二次定型 → 硫化 → 泄压 → 开模 → 卸胎 → （回待机）。
           待机相等 xStart 上升沿（必须边沿，防上电即在启动位自动合模）；
           装胎相给装胎命令等装胎到位反馈；合模相给合模命令等合模到位反馈；
           一次定型相开一次定型阀，等胶囊压力达 fShapePressKpa；二次定型相同理但压力窗更高；
           硫化相开主蒸汽阀，等 tCureS 且模温不低于 fCureTargetC − fTempBandK；
           泄压相开泄压阀，等压力降到 fVentPressKpa 以下；开模相等开模到位反馈；
           卸胎相等卸胎到位反馈，完成后置 xDone 锁存并回待机（保持到 xStart 撤下）。
        2) 每相独立超时 + 整序总超时：八个工作相各配「相定时 + 裕量」超时点，
           tonTotal 兜底整序总时长，九个超时源并发监视，任一命中即锁码进故障相。
        3) 硫化过程温度保护：硫化相内模温跌破 fCureTargetC − fTempBandK 即锁码 0337，
           这是欠硫的直接成因（温度不足则等效硫化时间按 Arrhenius 指数衰减）。
  边界条件：1) 非有限值闸：胶囊压力、模温、目标温度、压力阈、温度带宽、周期先过
           NOT(x > -DL_BIG AND x < DL_BIG)，同时拦 NaN 与 Inf；命中即锁码 0343 进故障相，
           绝不把 NaN 拿去与压力/温度阈比较（NaN 比较恒假会让放行条件永不成立，也永不报错，R19）。
        2) 周期入参闸（R21）：本件不做斜率运算，fCycleS 仅作观测与工艺记录；
           非法周期改用缺省 DL_CYCLE_DEF = 0.1 s，并在组态闸中一并锁码 0343（同码归因，内部成员分离）。
        3) 阈值域闸：0.0 < fShapePressKpa < fCurePressKpa、fVentPressKpa < fShapePressKpa、
           fTempBandK > DL_EPS，越域锁码 0343（定型压力窗倒置会让压力判据永不成立）。
        4) 单点赋值（R26）：九个命令位与 xDone / xBusy 全部在段 8 统一出口写一次，
           相位内只改 _eState 与锁存位，不在分支内各写一遍命令。
        5) 定时器周期刷新（R7）：十七个 TON 与两个边沿实例全部在 CASE 之外无条件调用，
           IN 由状态导出，相迁移即 IN 归假自复位（R188）。
        6) 故障解除路径：故障相内 xReset 上升沿 AND NOT xFault AND 入参/组态合法 → 清锁存回待机，
           回待机后必须重新给 xStart 上升沿才能再启动（不自恢复）。
        7) 状态机兜底：CASE 全态覆盖 + ELSE 强制回故障相并置码 0344、清全部输出。
        8) 输出安全初值（R25）：九个命令位初值 FALSE（失电即安全侧：不开阀不合模），
           xDone / xBusy 初值 FALSE，待机相显式赋值。
  量纲自证：fBladderPressKpa 与三个压力阈同为 [kPa]，比较合法；
           fMoldTempC / fCureTargetC 为 [degC]，fTempBandK 为温差不 [K]，degC 差值以 K 计，合法；
           所有时间引脚为 [TIME]，相超时点 = [TIME] + [TIME] = [TIME]，与 TON 的 PT 同量纲。
  码表 Error codes（本件子带 0091_033x / 034x，故障级一律 3 行内置 _uFault/_bFault/_eState）:
    16#0091_0331 信息级：装胎相等待装胎到位反馈（不置故障位）
    16#0091_0332 故障级：装胎相超时
    16#0091_0333 故障级：合模相超时（合模未到位）
    16#0091_0334 故障级：一次定型相超时（压力未达一次定型窗）
    16#0091_0335 故障级：二次定型相超时（压力未达二次定型窗）
    16#0091_0336 故障级：硫化相超时（等效硫化时间未跑完）
    16#0091_0337 故障级：硫化相模温低于下限（欠硫风险）
    16#0091_0338 故障级：泄压相超时（压力未泄尽）
    16#0091_0339 故障级：开模相超时（开模未到位）
    16#0091_0340 故障级：卸胎相超时（卸胎未到位）
    16#0091_0341 故障级：整序总超时
    16#0091_0342 故障级：外部故障输入 xFault
    16#0091_0343 故障级：入参非有限，或压力/温度/周期组态越域
    16#0091_0344 故障级：状态机落 ELSE 兜底（非法相位 ID）
    16#0091_0345 信息级：周期完成保持中，等待撤令（不置故障位）

  修订历史 Revision :
    2026-11-25  v1.0.0  R91 首版
*)

TYPE E_DL_TcsPressState :
(
    eTcsPressIdle   := 0,     // 待机：等启动上升沿，全命令撤销 / Idle, awaiting start, all commands dropped
    eTcsPressLoad   := 10,    // 装胎：给装胎命令等到位 / Loading, awaiting the load-done feedback
    eTcsPressClose  := 20,    // 合模：给合模命令等到位 / Closing, awaiting the closed feedback
    eTcsPressShape1 := 30,    // 一次定型：开一次定型阀等压力 / First shaping, awaiting the pressure window
    eTcsPressShape2 := 40,    // 二次定型：开二次定型阀等压力 / Second shaping, awaiting the pressure window
    eTcsPressCure   := 50,    // 硫化：开主蒸汽阀等时间与模温 / Curing, awaiting time and mold temperature
    eTcsPressVent   := 60,    // 泄压：开泄压阀等压力降 / Venting, awaiting the pressure drop
    eTcsPressOpen   := 70,    // 开模：给开模命令等到位 / Opening, awaiting the open feedback
    eTcsPressUnload := 80,    // 卸胎：给卸胎命令等到位 / Unloading, awaiting the unload-done feedback
    eTcsPressFault  := 90     // 故障：锁存待解除 / Fault, latched awaiting release
);
END_TYPE

FUNCTION_BLOCK FB_DL_TireCurePressSeq
VAR_INPUT
    xStart          : BOOL;    // 循环启动指令（上升沿有效）[bool] / Cycle start command, edge triggered [bool]
    xReset          : BOOL;    // 故障复位（上升沿有效）[bool] / Fault reset, rising edge [bool]
    xFault          : BOOL;    // 外部故障汇总 [bool] / External fault aggregate [bool]
    xLoadDoneFb     : BOOL;    // 装胎到位反馈 [bool] / Load-done feedback [bool]
    xClosedFb       : BOOL;    // 合模到位反馈 [bool] / Mold-closed feedback [bool]
    xOpenFb         : BOOL;    // 开模到位反馈 [bool] / Mold-open feedback [bool]
    xUnloadDoneFb   : BOOL;    // 卸胎到位反馈 [bool] / Unload-done feedback [bool]
    fBladderPressKpa : REAL;   // 胶囊实测压力 [kPa] / Measured bladder pressure [kPa]
    fMoldTempC      : REAL;    // 模温实测值 [degC] / Measured mold temperature [degC]
    fCureTargetC    : REAL;    // 硫化目标模温 [degC] / Curing target mold temperature [degC]
    fTempBandK      : REAL;    // 模温允许下偏带宽 [K] / Permitted mold temperature undershoot band [K]
    fShapePressKpa  : REAL;    // 定型压力窗（一次/二次共用下限）[kPa] / Shaping pressure window [kPa]
    fCurePressKpa   : REAL;    // 硫化压力窗（须高于定型窗）[kPa] / Curing pressure window [kPa]
    fVentPressKpa   : REAL;    // 泄压完成压力上限 [kPa] / Vent-complete pressure ceiling [kPa]
    fCycleS         : REAL;    // 任务周期（观测用）[s] / Task cycle time, for observation [s]
    tLoadS          : TIME;    // 装胎相设定时长 [TIME] / Loading phase duration [TIME]
    tCloseS         : TIME;    // 合模相设定时长 [TIME] / Closing phase duration [TIME]
    tShape1S        : TIME;    // 一次定型相设定时长 [TIME] / First shaping duration [TIME]
    tShape2S        : TIME;    // 二次定型相设定时长 [TIME] / Second shaping duration [TIME]
    tCureS          : TIME;    // 硫化相设定时长 [TIME] / Curing phase duration [TIME]
    tVentS          : TIME;    // 泄压相设定时长 [TIME] / Venting phase duration [TIME]
    tOpenS          : TIME;    // 开模相设定时长 [TIME] / Opening phase duration [TIME]
    tUnloadS        : TIME;    // 卸胎相设定时长 [TIME] / Unloading phase duration [TIME]
END_VAR
VAR_OUTPUT
    xLoadCmd        : BOOL;    // 装胎命令（安全侧：故障时停）[bool] / Load command, fail-safe [bool]
    xCloseCmd       : BOOL;    // 合模命令（安全侧：故障时停）[bool] / Close command, fail-safe [bool]
    xShape1ValveCmd : BOOL;    // 一次定型阀命令（安全侧：故障时关）[bool] / First shaping valve command [bool]
    xShape2ValveCmd : BOOL;    // 二次定型阀命令（安全侧：故障时关）[bool] / Second shaping valve command [bool]
    xCureSteamCmd   : BOOL;    // 硫化主蒸汽阀命令（安全侧：故障时关）[bool] / Curing steam valve command [bool]
    xVentValveCmd   : BOOL;    // 泄压阀命令（安全侧：故障时关）[bool] / Vent valve command [bool]
    xOpenCmd        : BOOL;    // 开模命令（安全侧：故障时停）[bool] / Open command, fail-safe [bool]
    xUnloadCmd      : BOOL;    // 卸胎命令（安全侧：故障时停）[bool] / Unload command, fail-safe [bool]
    xDone           : BOOL;    // 周期完成保持位 [bool] / Cycle complete held flag [bool]
    xBusy           : BOOL;    // 循环进行中 [bool] / Cycle busy [bool]
    eState          : E_DL_TcsPressState;   // 状态出口，段尾单点映射 / State outlet, single-point mapped
    nErrId          : UDINT;   // 事件码，0 = 无事件 / Event code, 0 = none
END_VAR
VAR
    tonLoad         : TON;     // 装胎相正常定时 [TIME] / Loading phase timer
    tonLoadOv       : TON;     // 装胎相超时定时 [TIME] / Loading phase overrun timer
    tonClose        : TON;     // 合模相正常定时 [TIME] / Closing phase timer
    tonCloseOv      : TON;     // 合模相超时定时 [TIME] / Closing phase overrun timer
    tonShape1       : TON;     // 一次定型相正常定时 [TIME] / First shaping phase timer
    tonShape1Ov     : TON;     // 一次定型相超时定时 [TIME] / First shaping phase overrun timer
    tonShape2       : TON;     // 二次定型相正常定时 [TIME] / Second shaping phase timer
    tonShape2Ov     : TON;     // 二次定型相超时定时 [TIME] / Second shaping phase overrun timer
    tonCure         : TON;     // 硫化相正常定时 [TIME] / Curing phase timer
    tonCureOv       : TON;     // 硫化相超时定时 [TIME] / Curing phase overrun timer
    tonVent         : TON;     // 泄压相正常定时 [TIME] / Venting phase timer
    tonVentOv       : TON;     // 泄压相超时定时 [TIME] / Venting phase overrun timer
    tonOpen         : TON;     // 开模相正常定时 [TIME] / Opening phase timer
    tonOpenOv       : TON;     // 开模相超时定时 [TIME] / Opening phase overrun timer
    tonUnload       : TON;     // 卸胎相正常定时 [TIME] / Unloading phase timer
    tonUnloadOv     : TON;     // 卸胎相超时定时 [TIME] / Unloading phase overrun timer
    tonTotal        : TON;     // 整序总超时定时 [TIME] / Whole-sequence total timeout timer
    rtStart         : R_TRIG;  // 启动上升沿检测 [bool] / Start rising edge detector
    rtReset         : R_TRIG;  // 复位上升沿检测 [bool] / Reset rising edge detector
    _eState         : E_DL_TcsPressState := E_DL_TcsPressState.eTcsPressIdle;   // 内部相位（CASE 唯一写入目标）
    _eStatePrev     : E_DL_TcsPressState := E_DL_TcsPressState.eTcsPressIdle;   // 上一拍相位快照（周期末更新）
    _fCycleUseS     : REAL := 0.1;    // 实际使用的周期值 [s] / Cycle time actually used [s]
    _fTempLowK      : REAL := 0.0;    // 硫化模温下限 [degC] / Curing mold temperature low limit [degC]
    _fTempDevK      : REAL := 0.0;    // 模温低于目标的下偏量 [K] / Mold temperature undershoot [K]
    _bFinOk         : BOOL := FALSE;  // 实值入参有限性总闸结果 / Finiteness gate aggregate result
    _bCfgOk         : BOOL := FALSE;  // 压力/温度/周期组态域闸结果 / Configuration domain gate result
    _bActive        : BOOL := FALSE;  // 序激活（装胎至卸胎八相之一）[bool] / Sequence active flag
    _bDoneL         : BOOL := FALSE;  // 完成位锁存（跨相保持）[bool] / Done latch held across phases
    _bFault         : BOOL := FALSE;  // 故障锁存位 [bool] / Latched fault flag
    _iPhaseChg      : INT := 0;       // 本拍相位切换计数（观测用）[-] / Phase-change count this cycle [-]
    _uInfo          : UDINT := 16#0000_0000;   // 信息码，每拍重算 / Info code, recomputed every cycle
    _uFault         : UDINT := 16#0000_0000;   // 故障码锁存 / Latched fault code
END_VAR
VAR CONSTANT
    DL_EPS          : REAL := 1.0E-9;     // 数值零闸阈值 [-] / Numeric zero gate threshold [-]
    DL_BIG          : REAL := 1.0E12;     // 非有限值闸量级上限 [-] / Finiteness gate magnitude [-]
    DL_CYCLE_DEF    : REAL := 0.1;        // 缺省任务周期 [s] / Default task cycle time [s]
    DL_CYCLE_MIN    : REAL := 0.001;      // 周期合理下限 [s] / Cycle time reasonable low bound [s]
    DL_CYCLE_MAX    : REAL := 10.0;       // 周期合理上限 [s] / Cycle time reasonable high bound [s]
    DL_PRESS_HI     : REAL := 10000.0;    // 压力量级闸上限 [kPa] / Pressure magnitude upper bound [kPa]
    DL_T_SPAN       : REAL := 500.0;      // 温度量级闸跨度 [degC] / Temperature magnitude gate span [degC]
    DL_OVER_MARGIN  : TIME := T#30S;      // 相超时相对正常定时的裕量 [TIME] / Phase overrun margin [TIME]
    DL_TOTAL_MAX    : TIME := T#4H;       // 整序总超时上限 [TIME] / Whole-sequence total timeout [TIME]
END_VAR

(* —— 段 0：单拍量预清零（锁存量 _uFault/_bFault/_bDoneL/_eStatePrev 不入清单，R187①） —— *)
_uInfo := 16#0000_0000;                     // 信息码每拍重算 / Info code recomputed
_iPhaseChg := 0;                            // 相位切换计数每拍重算 / Phase-change counter recomputed
nErrId := 16#0000_0000;                     // 事件码缺省无事件 / Event code defaults to none

(* —— 段 1：非有限值闸与组态域闸（R19：不拿 NaN 去比较压力与温度阈） —— *)
_bFinOk := (fBladderPressKpa > -DL_BIG) AND (fBladderPressKpa < DL_BIG)
           AND (fMoldTempC > -DL_BIG) AND (fMoldTempC < DL_BIG)
           AND (fCureTargetC > -DL_BIG) AND (fCureTargetC < DL_BIG)
           AND (fTempBandK > -DL_BIG) AND (fTempBandK < DL_BIG)
           AND (fShapePressKpa > -DL_BIG) AND (fShapePressKpa < DL_BIG)
           AND (fCurePressKpa > -DL_BIG) AND (fCurePressKpa < DL_BIG)
           AND (fVentPressKpa > -DL_BIG) AND (fVentPressKpa < DL_BIG)
           AND (fCycleS > -DL_BIG) AND (fCycleS < DL_BIG);
_bCfgOk := (fVentPressKpa >= 0.0)                          // 泄压上限不得为负
           AND (fShapePressKpa > fVentPressKpa)            // 定型窗必须高于泄压窗
           AND (fCurePressKpa > fShapePressKpa)            // 硫化窗必须高于定型窗（压力窗单调）
           AND (fCurePressKpa <= DL_PRESS_HI)              // 硫化窗须在压力量级内
           AND (fTempBandK > DL_EPS)                       // 温度带宽必须为正
           AND (ABS(fCureTargetC) <= DL_T_SPAN)            // 目标模温量级闸
           AND (ABS(fMoldTempC) <= DL_T_SPAN)              // 实测模温量级闸
           AND (fCycleS >= DL_CYCLE_MIN) AND (fCycleS <= DL_CYCLE_MAX);

IF _bCfgOk THEN
    _fCycleUseS := fCycleS;                 // 合法周期原值使用（本件仅观测用）
ELSE
    _fCycleUseS := DL_CYCLE_DEF;            // 非法周期一律用缺省 0.1 s
END_IF

(* —— 段 2：派生态（序激活、模温下偏量） —— *)
_bActive := (_eState = E_DL_TcsPressState.eTcsPressLoad)
            OR (_eState = E_DL_TcsPressState.eTcsPressClose)
            OR (_eState = E_DL_TcsPressState.eTcsPressShape1)
            OR (_eState = E_DL_TcsPressState.eTcsPressShape2)
            OR (_eState = E_DL_TcsPressState.eTcsPressCure)
            OR (_eState = E_DL_TcsPressState.eTcsPressVent)
            OR (_eState = E_DL_TcsPressState.eTcsPressOpen)
            OR (_eState = E_DL_TcsPressState.eTcsPressUnload);
_fTempLowK := fCureTargetC - fTempBandK;                                  // 硫化模温下限 [degC]
_fTempDevK := fCureTargetC - fMoldTempC;                                  // 模温下偏量 [K]

(* —— 段 3：定时器与边沿无条件周期刷新（R7：调用语句不得置于 IF/CASE 内） —— *)
rtStart(CLK := xStart);                                                                    // 启动上升沿，每拍必调
rtReset(CLK := xReset);                                                                    // 复位上升沿，每拍必调
tonLoad(IN := (_eState = E_DL_TcsPressState.eTcsPressLoad), PT := tLoadS);                 // 装胎相正常定时
tonLoadOv(IN := (_eState = E_DL_TcsPressState.eTcsPressLoad), PT := tLoadS + DL_OVER_MARGIN);         // 装胎超时点
tonClose(IN := (_eState = E_DL_TcsPressState.eTcsPressClose), PT := tCloseS);              // 合模相正常定时
tonCloseOv(IN := (_eState = E_DL_TcsPressState.eTcsPressClose), PT := tCloseS + DL_OVER_MARGIN);       // 合模超时点
tonShape1(IN := (_eState = E_DL_TcsPressState.eTcsPressShape1), PT := tShape1S);           // 一次定型正常定时
tonShape1Ov(IN := (_eState = E_DL_TcsPressState.eTcsPressShape1), PT := tShape1S + DL_OVER_MARGIN);    // 一次定型超时点
tonShape2(IN := (_eState = E_DL_TcsPressState.eTcsPressShape2), PT := tShape2S);           // 二次定型正常定时
tonShape2Ov(IN := (_eState = E_DL_TcsPressState.eTcsPressShape2), PT := tShape2S + DL_OVER_MARGIN);    // 二次定型超时点
tonCure(IN := (_eState = E_DL_TcsPressState.eTcsPressCure), PT := tCureS);                 // 硫化相正常定时
tonCureOv(IN := (_eState = E_DL_TcsPressState.eTcsPressCure), PT := tCureS + DL_OVER_MARGIN);          // 硫化超时点
tonVent(IN := (_eState = E_DL_TcsPressState.eTcsPressVent), PT := tVentS);                 // 泄压相正常定时
tonVentOv(IN := (_eState = E_DL_TcsPressState.eTcsPressVent), PT := tVentS + DL_OVER_MARGIN);          // 泄压超时点
tonOpen(IN := (_eState = E_DL_TcsPressState.eTcsPressOpen), PT := tOpenS);                 // 开模相正常定时
tonOpenOv(IN := (_eState = E_DL_TcsPressState.eTcsPressOpen), PT := tOpenS + DL_OVER_MARGIN);          // 开模超时点
tonUnload(IN := (_eState = E_DL_TcsPressState.eTcsPressUnload), PT := tUnloadS);           // 卸胎相正常定时
tonUnloadOv(IN := (_eState = E_DL_TcsPressState.eTcsPressUnload), PT := tUnloadS + DL_OVER_MARGIN);    // 卸胎超时点
tonTotal(IN := _bActive, PT := DL_TOTAL_MAX);                                              // 整序总超时

(* —— 段 4：全局故障拦截（优先级最高；已锁存则不再改写码值，禁同拍抹除） —— *)
IF xFault AND (NOT _bFault) THEN
    _uFault := 16#0091_0342;                // 故障级：外部故障输入
    _bFault := TRUE;                        // 锁存（3 行内置，R45 配对）
    _eState := E_DL_TcsPressState.eTcsPressFault;
END_IF
IF ((NOT _bFinOk) OR (NOT _bCfgOk)) AND (NOT _bFault) THEN
    _uFault := 16#0091_0343;                // 故障级：入参非有限或组态越域（内部成员已分离）
    _bFault := TRUE;                        // 锁存
    _eState := E_DL_TcsPressState.eTcsPressFault;
END_IF
IF tonTotal.Q AND _bActive AND (NOT _bFault) THEN
    _uFault := 16#0091_0341;                // 故障级：整序总超时
    _bFault := TRUE;                        // 锁存
    _eState := E_DL_TcsPressState.eTcsPressFault;
END_IF
IF (_eState = E_DL_TcsPressState.eTcsPressCure)
   AND (_fTempDevK > fTempBandK) AND (NOT _bFault) THEN
    _uFault := 16#0091_0337;                // 故障级：硫化模温低于下限（欠硫风险）
    _bFault := TRUE;                        // 锁存
    _eState := E_DL_TcsPressState.eTcsPressFault;
END_IF

(* —— 段 5：相位机（只做迁移；出口在段 7 单点映射） —— *)
CASE _eState OF

E_DL_TcsPressState.eTcsPressIdle:
    IF NOT xStart THEN
        _bDoneL := FALSE;                   // 撤令即清完成位，为下一模重新武装
    ELSIF rtStart.Q THEN
        _bDoneL := FALSE;                   // 新循环开始：清完成位（迁移前一次性清）
        _eState := E_DL_TcsPressState.eTcsPressLoad;          // 进装胎相
    END_IF

E_DL_TcsPressState.eTcsPressLoad:
    IF tonLoadOv.Q THEN
        _uFault := 16#0091_0332;            // 故障级：装胎相超时
        _bFault := TRUE;                    // 锁存
        _eState := E_DL_TcsPressState.eTcsPressFault;
    ELSIF tonLoad.Q AND xLoadDoneFb THEN
        _eState := E_DL_TcsPressState.eTcsPressClose;         // 本拍合法事件优先于超时迁移（R275）
    ELSE
        _uInfo := 16#0091_0331;             // 信息级：等装胎到位反馈（不置故障位）
    END_IF

E_DL_TcsPressState.eTcsPressClose:
    IF tonCloseOv.Q THEN
        _uFault := 16#0091_0333;            // 故障级：合模相超时
        _bFault := TRUE;                    // 锁存
        _eState := E_DL_TcsPressState.eTcsPressFault;
    ELSIF xClosedFb THEN
        _eState := E_DL_TcsPressState.eTcsPressShape1;        // 合模到位：进一次定型相
    END_IF

E_DL_TcsPressState.eTcsPressShape1:
    IF tonShape1Ov.Q THEN
        _uFault := 16#0091_0334;            // 故障级：一次定型相超时
        _bFault := TRUE;                    // 锁存
        _eState := E_DL_TcsPressState.eTcsPressFault;
    ELSIF (fBladderPressKpa >= fShapePressKpa) AND tonShape1.Q THEN
        _eState := E_DL_TcsPressState.eTcsPressShape2;        // 压力窗达成：进二次定型相
    END_IF

E_DL_TcsPressState.eTcsPressShape2:
    IF tonShape2Ov.Q THEN
        _uFault := 16#0091_0335;            // 故障级：二次定型相超时
        _bFault := TRUE;                    // 锁存
        _eState := E_DL_TcsPressState.eTcsPressFault;
    ELSIF (fBladderPressKpa >= fCurePressKpa) AND tonShape2.Q THEN
        _eState := E_DL_TcsPressState.eTcsPressCure;          // 压力窗达成：进硫化相
    END_IF

E_DL_TcsPressState.eTcsPressCure:
    IF tonCureOv.Q THEN
        _uFault := 16#0091_0336;            // 故障级：硫化相超时
        _bFault := TRUE;                    // 锁存
        _eState := E_DL_TcsPressState.eTcsPressFault;
    ELSIF tonCure.Q THEN
        _eState := E_DL_TcsPressState.eTcsPressVent;          // 等效硫化时间到：进泄压相
    END_IF

E_DL_TcsPressState.eTcsPressVent:
    IF tonVentOv.Q THEN
        _uFault := 16#0091_0338;            // 故障级：泄压相超时
        _bFault := TRUE;                    // 锁存
        _eState := E_DL_TcsPressState.eTcsPressFault;
    ELSIF (fBladderPressKpa <= fVentPressKpa) AND tonVent.Q THEN
        _eState := E_DL_TcsPressState.eTcsPressOpen;          // 压力泄尽：进开模相
    END_IF

E_DL_TcsPressState.eTcsPressOpen:
    IF tonOpenOv.Q THEN
        _uFault := 16#0091_0339;            // 故障级：开模相超时
        _bFault := TRUE;                    // 锁存
        _eState := E_DL_TcsPressState.eTcsPressFault;
    ELSIF xOpenFb AND tonOpen.Q THEN
        _eState := E_DL_TcsPressState.eTcsPressUnload;        // 开模到位：进卸胎相
    END_IF

E_DL_TcsPressState.eTcsPressUnload:
    IF tonUnloadOv.Q THEN
        _uFault := 16#0091_0340;            // 故障级：卸胎相超时
        _bFault := TRUE;                    // 锁存
        _eState := E_DL_TcsPressState.eTcsPressFault;
    ELSIF xUnloadDoneFb AND tonUnload.Q THEN
        _bDoneL := TRUE;                    // 完成位锁存（跨相保持，段 7 单点映射）
        _eState := E_DL_TcsPressState.eTcsPressIdle;          // 回待机，完成位保持到撤令
    END_IF

E_DL_TcsPressState.eTcsPressFault:
    IF rtReset.Q AND (NOT xFault) AND _bFinOk AND _bCfgOk THEN
        _bFault := FALSE;                   // 解除路径：复位沿 + 外部故障消失 + 入参/组态合法（可达，R188）
        _uFault := 16#0000_0000;            // 清锁存码
        _bDoneL := FALSE;                   // 完成位一并清，避免故障后误报完成
        _eState := E_DL_TcsPressState.eTcsPressIdle;          // 回待机，需新上升沿才可再启动
    END_IF

ELSE
    _uFault := 16#0091_0344;                // 故障级：非法相位 ID 兜底
    _bFault := TRUE;                        // 锁存
    _bDoneL := FALSE;                       // 完成位清
    _eState := E_DL_TcsPressState.eTcsPressFault;             // 强制回故障相

END_CASE

(* —— 段 6：后置段（相位快照在迁移判断之后统一更新） —— *)
IF _eState <> _eStatePrev THEN
    _iPhaseChg := _iPhaseChg + 1;           // 相位已切换：记一拍切换事件（观测用）
END_IF
_eStatePrev := _eState;                     // 快照在周期末尾统一更新

(* —— 段 7：出口单点映射（名实同源；九个命令位由状态导出，故障侧一律撤销） —— *)
xLoadCmd := (_eState = E_DL_TcsPressState.eTcsPressLoad) AND (NOT _bFault);               // 装胎命令
xCloseCmd := (_eState = E_DL_TcsPressState.eTcsPressClose) AND (NOT _bFault);             // 合模命令
xShape1ValveCmd := (_eState = E_DL_TcsPressState.eTcsPressShape1) AND (NOT _bFault);      // 一次定型阀
xShape2ValveCmd := (_eState = E_DL_TcsPressState.eTcsPressShape2) AND (NOT _bFault);      // 二次定型阀
xCureSteamCmd := (_eState = E_DL_TcsPressState.eTcsPressCure) AND (NOT _bFault);          // 硫化蒸汽阀
xVentValveCmd := (_eState = E_DL_TcsPressState.eTcsPressVent) AND (NOT _bFault);          // 泄压阀
xOpenCmd := (_eState = E_DL_TcsPressState.eTcsPressOpen) AND (NOT _bFault);               // 开模命令
xUnloadCmd := (_eState = E_DL_TcsPressState.eTcsPressUnload) AND (NOT _bFault);           // 卸胎命令
xDone := _bDoneL AND (NOT _bFault);                                                       // 完成位出口
xBusy := _bActive AND (NOT _bFault);                                                      // 进行中出口
eState := _eState;                                                                        // 状态出口单点映射
IF _bFault THEN
    nErrId := _uFault;                      // 故障锁存码回放（不在故障相按当下输入重推断）
ELSIF _bDoneL THEN
    nErrId := 16#0091_0345;                 // 信息级：周期完成保持中，等待撤令
ELSE
    nErrId := _uInfo;                       // 信息码
END_IF

END_FUNCTION_BLOCK

(* ---- FB_DL_TobaccoCuttingLineSeq.st ---- *)
(*
 * FB_DL_TobaccoCuttingLineSeq | C4 | DL_Process
 * 功能：制丝线「进料→切丝→烘丝→冷却→掺配→完成」工段序列控制；每相独立使能出口 + 独立 TON 超时，超时/参数非法一律回 FAULT 并撤销全部命令       单位：水分 [%]、rTimeoutS [s]、nFaultCode [INT 码位]
 * 工况边界：出口水分 rMoistOutPct 与目标 rMoistTargetPct 须在 0~100 % 且有限，DRYING 只在 |出口−目标|≤0.5 % 时转 COOLING；rTimeoutS 须 >0；xStart 为电平输入但只用上升沿启动（停车后须先撤 xStart 再给，防自恢复）；xStop 在任意相生效，按逆序（先切丝/烘丝，后进料）在同拍归零全部命令，物理减速由变频器斜坡完成；xComplete 为 DONE 相状态量（非单拍脉冲），下游取上升沿
 * 代数值回代：rMoistOutPct=12.0、rMoistTargetPct=12.0 → |Δ|=0 ≤0.5 满足转 COOLING；rMoistOutPct=13.2 → |Δ|=1.2 >0.5 驻留 DRYING 直至 9401（spec 判定式一致）
 * 开源溯源：clean-room 自研，未复制任何第三方代码（无外部来源）
 *)
(*
 * 码位总账（本件故障码全清单，逐条在实现分支中可到达；故障级锁存回放）：
 * 9401 烘丝水分偏差超时 / 9402 进料超时或进料未就绪 / 9403 切丝超时或切丝未就绪 / 9404 冷却相输送就绪丢失 / 9406 水分越界或状态机兜底（故障锁存，清除沿 = xStart 下降沿）；9405 本件预留未使用——掺配相以驻留定时正常完成，无独立故障判据，故不设该码位（码表与实现逐分支对齐）
 *)

TYPE E_DL_TobCutPhase :
(
    IDLE    := 0,       // 待机，全部命令撤销 | idle, every command withdrawn
    FEEDING := 10,      // 进料相，仅进料命令 | feeding phase, feed command only
    CUTTING := 20,      // 切丝相，进料 + 切丝命令 | cutting phase, feed plus cutter
    DRYING  := 30,      // 烘丝相，进料 + 切丝 + 烘丝命令 | drying phase, feed plus cutter plus dryer
    COOLING := 40,      // 冷却相，仅输送风机（进料）命令 | cooling phase, conveying command only
    BLENDING:= 50,      // 掺配相，仅掺配命令 | blending phase, blending command only
    DONE    := 60,      // 完成相，全部命令撤销，xComplete 置位 | done phase, all commands withdrawn, xComplete raised
    FAULT   := 90       // 故障相，全部命令强制 FALSE，码位锁存 | fault phase, all commands forced FALSE, the code is latched
);
END_TYPE

FUNCTION_BLOCK FB_DL_TobaccoCuttingLineSeq
VAR_INPUT
    xStart          : BOOL;          // 启动（下降沿兼作故障复位沿）| start, its falling edge also resets a latched fault
    xStop           : BOOL;          // 停止（任意相生效，逆序停车）| stop, effective in any phase and stopping in reverse order
    xFeedReady      : BOOL;          // 进料段就绪 | feeding section ready
    xCutterReady    : BOOL;          // 切丝机就绪 | cutter ready
    xDryerReady     : BOOL;          // 烘丝机就绪 | dryer ready
    rMoistOutPct    : REAL;          // 烘丝出口水分 | dryer outlet moisture [%]
    rMoistTargetPct : REAL := 12.0;  // 烘丝出口目标水分 | dryer outlet moisture target [%]
    rTimeoutS       : REAL := 60.0;  // 每相超时设定 | per-phase timeout setting [s]
END_VAR
VAR_OUTPUT
    xFeedCmd   : BOOL;               // 进料/输送命令（FEEDING/CUTTING/DRYING/COOLING 相独立使能）| feed command, independent enable of those phases
    xCutterCmd : BOOL;               // 切丝命令（CUTTING/DRYING 相独立使能）| cutter command, independent enable of those phases
    xDryerCmd  : BOOL;               // 烘丝命令（DRYING 相独立使能）| dryer command, independent enable of DRYING
    xBlendCmd  : BOOL;               // 掺配命令（BLENDING 相独立使能）| blending command, independent enable of BLENDING
    ePhase     : E_DL_TobCutPhase;   // 当前相 | current phase
    xComplete  : BOOL;               // 完成状态量（DONE 相为 TRUE，非单拍脉冲）| completion level, true in DONE
    xFault     : BOOL;               // 故障标志 | fault flag
    nFaultCode : INT;                // 故障码，锁存至复位沿 | fault code latched until the reset edge
END_VAR
VAR
    tonFeed  : TON;                  // FEEDING 相超时定时器 | timeout of the FEEDING phase
    tonCut   : TON;                  // CUTTING 相超时定时器 | timeout of the CUTTING phase
    tonDry   : TON;                  // DRYING 相超时定时器 | timeout of the DRYING phase
    tonCool  : TON;                  // COOLING 相超时定时器 | timeout of the COOLING phase
    tonBlend : TON;                  // BLENDING 相超时定时器 | timeout of the BLENDING phase
    tonDone  : TON;                  // DONE 相驻留定时器 | dwell timer of the DONE phase
    fbStartFall : F_TRIG;            // xStart 下降沿（故障复位沿）| falling edge of xStart, the fault reset edge
    fbStartRise : R_TRIG;            // xStart 上升沿（唯一启动沿，防止停车后自动重启）| rising edge of xStart, the single start edge preventing an auto restart
    xParamOk : BOOL;                 // 超时参数合法 | timeout parameter is legal
    xFinMoist: BOOL;                 // 出口水分有限性 | outlet moisture is finite
    xMoistBad: BOOL;                 // 出口水分越界或非有限 | outlet moisture out of range or non-finite
    xInBand  : BOOL;                 // 水分落在目标 ±0.5 % 容带内 | moisture inside the target band
    nTmoMs   : UDINT := 60000;       // 超时毫秒数（缺省值防首拍 PT=0 假超时）| timeout in milliseconds, default prevents a zero PT on the first scan
    nCodeLatch : INT;                // 故障码锁存副本 | latched copy of the fault code
END_VAR
VAR CONSTANT
    DL_TCS_BAND_PCT : REAL := 0.5;   // 水分容带半宽 | moisture band half width [%]
    DL_TCS_PCT_MIN  : REAL := 0.0;   // 水分下限 | lower moisture limit [%]
    DL_TCS_PCT_MAX  : REAL := 100.0; // 水分上限 | upper moisture limit [%]
    DL_TCS_C_MOIST  : INT := 9401;   // 烘丝水分偏差超时 | drying moisture deviation timeout
    DL_TCS_C_FEED   : INT := 9402;   // 进料超时/未就绪 | feeding timeout or not ready
    DL_TCS_C_CUT    : INT := 9403;   // 切丝超时/未就绪 | cutting timeout or not ready
    DL_TCS_C_COOL   : INT := 9404;   // 冷却超时 | cooling timeout
    DL_TCS_C_BAD    : INT := 9406;   // 水分越界或兜底 | moisture out of range or fallback
END_VAR

// 段1｜参数与采样门禁（先判后用：REAL→UDINT 换算在闸后进行，结果供段2 定时器使用）
xParamOk := (rTimeoutS = rTimeoutS) AND ((rTimeoutS - rTimeoutS) = 0.0) AND (rTimeoutS > 0.0);
IF xParamOk THEN
    nTmoMs := REAL_TO_UDINT(rTimeoutS * 1000.0);
ELSE
    nTmoMs := 60000;                 // 参数非法时取保守超时 | conservative timeout when the parameter is illegal
END_IF
xFinMoist := (rMoistOutPct = rMoistOutPct) AND ((rMoistOutPct - rMoistOutPct) = 0.0)
             AND (rMoistTargetPct = rMoistTargetPct) AND ((rMoistTargetPct - rMoistTargetPct) = 0.0);
xMoistBad := (NOT xFinMoist)
             OR (rMoistOutPct < DL_TCS_PCT_MIN) OR (rMoistOutPct > DL_TCS_PCT_MAX)
             OR (rMoistTargetPct < DL_TCS_PCT_MIN) OR (rMoistTargetPct > DL_TCS_PCT_MAX);
xInBand := (NOT xMoistBad) AND (ABS(rMoistOutPct - rMoistTargetPct) <= DL_TCS_BAND_PCT);

// 段2｜六只定时器 + 两只边沿实例无条件周期刷新（R7，一相一只实例不跨相复用；PT 取自段1 已换算毫秒值）
tonFeed(IN := ePhase = E_DL_TobCutPhase.FEEDING, PT := UDINT_TO_TIME(nTmoMs));
tonCut(IN := ePhase = E_DL_TobCutPhase.CUTTING, PT := UDINT_TO_TIME(nTmoMs));
tonDry(IN := ePhase = E_DL_TobCutPhase.DRYING, PT := UDINT_TO_TIME(nTmoMs));
tonCool(IN := ePhase = E_DL_TobCutPhase.COOLING, PT := UDINT_TO_TIME(nTmoMs));
tonBlend(IN := ePhase = E_DL_TobCutPhase.BLENDING, PT := UDINT_TO_TIME(nTmoMs));
tonDone(IN := ePhase = E_DL_TobCutPhase.DONE, PT := UDINT_TO_TIME(nTmoMs));
fbStartFall(CLK := xStart);
fbStartRise(CLK := xStart);

// 段3｜输出预置（唯一预置点；CASE 内只置位，其后不再无条件清零）
xFeedCmd := FALSE;
xCutterCmd := FALSE;
xDryerCmd := FALSE;
xBlendCmd := FALSE;
xComplete := FALSE;
xFault := FALSE;
nFaultCode := 0;

// 段4｜全局闸：参数/水分非法 → 直接锁故障；xStop → 逆序停车并撤销全部命令
IF (NOT xParamOk) OR xMoistBad THEN
    nCodeLatch := DL_TCS_C_BAD;
    xFault := TRUE;
    nFaultCode := DL_TCS_C_BAD;
    xFeedCmd := FALSE;               // 逆序停车：下游先停 | reverse stop, downstream first
    xCutterCmd := FALSE;
    xDryerCmd := FALSE;
    xBlendCmd := FALSE;
    ePhase := E_DL_TobCutPhase.FAULT;
ELSIF xStop AND (ePhase <> E_DL_TobCutPhase.IDLE) THEN
    xCutterCmd := FALSE;             // 逆序停车第 1 步：切丝与烘丝先停 | reverse stop step 1, cutter and dryer first
    xDryerCmd := FALSE;
    xBlendCmd := FALSE;
    xFeedCmd := FALSE;               // 逆序停车第 2 步：进料后停（同拍置假，斜坡由变频器完成）| step 2, feed last
    ePhase := E_DL_TobCutPhase.IDLE;
END_IF

// 段5｜主状态机（ENUM + CASE，ELSE 兜底）
IF ePhase <> E_DL_TobCutPhase.FAULT THEN
CASE ePhase OF
E_DL_TobCutPhase.IDLE:
    // 拍 N：待机，无命令；仅 xStart 上升沿且进料就绪、无停车请求时启动（防停车后自恢复）
    IF fbStartRise.Q AND xFeedReady AND (NOT xStop) THEN
        ePhase := E_DL_TobCutPhase.FEEDING;      // 本拍行为：进料相（命令下拍由段6给出）| enter feeding
    END_IF

E_DL_TobCutPhase.FEEDING:
    // 拍 N：进料中，等切丝机就绪
    IF (NOT xFeedReady) THEN
        nCodeLatch := DL_TCS_C_FEED;             // 进料就绪丢失 | feed readiness lost
        xFault := TRUE;
        nFaultCode := DL_TCS_C_FEED;
        ePhase := E_DL_TobCutPhase.FAULT;
    ELSIF xCutterReady THEN
        ePhase := E_DL_TobCutPhase.CUTTING;      // 本拍行为：切丝机就绪转切丝 | cutter ready, enter cutting
    ELSIF tonFeed.Q THEN
        nCodeLatch := DL_TCS_C_FEED;             // 进料超时 | feeding timeout
        xFault := TRUE;
        nFaultCode := DL_TCS_C_FEED;
        ePhase := E_DL_TobCutPhase.FAULT;
    END_IF

E_DL_TobCutPhase.CUTTING:
    // 拍 N：切丝中，等烘丝机就绪
    IF NOT xCutterReady THEN
        nCodeLatch := DL_TCS_C_CUT;              // 切丝机就绪丢失 | cutter readiness lost
        xFault := TRUE;
        nFaultCode := DL_TCS_C_CUT;
        ePhase := E_DL_TobCutPhase.FAULT;
    ELSIF xDryerReady THEN
        ePhase := E_DL_TobCutPhase.DRYING;       // 本拍行为：烘丝机就绪转烘丝 | dryer ready, enter drying
    ELSIF tonCut.Q THEN
        nCodeLatch := DL_TCS_C_CUT;              // 切丝超时 | cutting timeout
        xFault := TRUE;
        nFaultCode := DL_TCS_C_CUT;
        ePhase := E_DL_TobCutPhase.FAULT;
    END_IF

E_DL_TobCutPhase.DRYING:
    // 拍 N：烘丝中，出口水分进入目标容带才转 COOLING
    IF NOT xDryerReady THEN
        nCodeLatch := DL_TCS_C_BAD;              // 烘丝机异常：按参数级故障处理 | dryer abnormality handled as a parameter-class fault
        xFault := TRUE;
        nFaultCode := DL_TCS_C_BAD;
        ePhase := E_DL_TobCutPhase.FAULT;
    ELSIF xInBand THEN
        ePhase := E_DL_TobCutPhase.COOLING;      // 本拍行为：水分达标转冷却 | moisture in band, enter cooling
    ELSIF tonDry.Q THEN
        nCodeLatch := DL_TCS_C_MOIST;            // 水分偏差超时：停在上限不转相 | moisture deviation timeout, hold the upper limit
        xFault := TRUE;
        nFaultCode := DL_TCS_C_MOIST;
        ePhase := E_DL_TobCutPhase.FAULT;
    END_IF

E_DL_TobCutPhase.COOLING:
    // 拍 N：冷却输送（输送机由进料段驱动），输送就绪丢失即报 9404；正常由驻留定时转掺配
    IF NOT xFeedReady THEN
        nCodeLatch := DL_TCS_C_COOL;                 // 冷却输送中断 | cooling conveying interrupted
        xFault := TRUE;
        nFaultCode := DL_TCS_C_COOL;
        ePhase := E_DL_TobCutPhase.FAULT;
    ELSIF tonCool.Q THEN
        ePhase := E_DL_TobCutPhase.BLENDING;         // 本拍行为：冷却完成转掺配 | cooling done, enter blending
    END_IF

E_DL_TobCutPhase.BLENDING:
    // 拍 N：掺配中，等掺配时间走完（驻留定时到即视为正常完成，不设故障码位，见头注释 9405 预留说明）
    IF tonBlend.Q THEN
        ePhase := E_DL_TobCutPhase.DONE;         // 本拍行为：掺配完成 | blending done
    END_IF

E_DL_TobCutPhase.DONE:
    // 拍 N：完成相，xComplete 由段6置位，驻留一个超时窗后回待机
    IF tonDone.Q OR (NOT xStart) THEN
        ePhase := E_DL_TobCutPhase.IDLE;         // 本拍行为：回待机 | back to idle
    END_IF

E_DL_TobCutPhase.FAULT:
    // 故障相（本段被外层 IF 排除，保留分支以满足穷举）
    xFault := TRUE;
    nFaultCode := nCodeLatch;

ELSE
    // 非法状态兜底：绝不停在未知相
    nCodeLatch := DL_TCS_C_BAD;
    xFault := TRUE;
    nFaultCode := DL_TCS_C_BAD;
    ePhase := E_DL_TobCutPhase.FAULT;
END_CASE
END_IF

// 段6｜每相独立使能出口（FAULT/IDLE/DONE 不置任何命令，天然强制 FALSE）
CASE ePhase OF
E_DL_TobCutPhase.FEEDING:
    xFeedCmd := TRUE;                        // 进料相独立使能出口 | independent enable of FEEDING
E_DL_TobCutPhase.CUTTING:
    xFeedCmd := TRUE;                        // 切丝相：进料保持 | cutting, keep feeding
    xCutterCmd := TRUE;                      // 切丝相独立使能出口 | independent enable of CUTTING
E_DL_TobCutPhase.DRYING:
    xFeedCmd := TRUE;                        // 烘丝相：进料保持 | drying, keep feeding
    xCutterCmd := TRUE;                      // 烘丝相：切丝保持 | drying, keep cutting
    xDryerCmd := TRUE;                       // 烘丝相独立使能出口 | independent enable of DRYING
E_DL_TobCutPhase.COOLING:
    xFeedCmd := TRUE;                        // 冷却相独立使能出口（输送风机）| independent enable of COOLING
E_DL_TobCutPhase.BLENDING:
    xBlendCmd := TRUE;                       // 掺配相独立使能出口 | independent enable of BLENDING
E_DL_TobCutPhase.DONE:
    xComplete := TRUE;                       // 完成状态量 | completion level
ELSE
    xFeedCmd := FALSE;                       // 其余相（含 FAULT）：命令强制 FALSE | all other phases force FALSE
    xCutterCmd := FALSE;
    xDryerCmd := FALSE;
    xBlendCmd := FALSE;
END_CASE

// 段7｜故障相锁存回放 + 复位沿（xStart 下降沿清除）
IF ePhase = E_DL_TobCutPhase.FAULT THEN
    xFault := TRUE;
    nFaultCode := nCodeLatch;                // 锁存回放，不按当下输入重推断 | republish the latch
    xFeedCmd := FALSE;
    xCutterCmd := FALSE;
    xDryerCmd := FALSE;
    xBlendCmd := FALSE;
    xComplete := FALSE;
    IF fbStartFall.Q THEN
        nCodeLatch := 0;                     // 清除边：xStart 下降沿（头注释已声明）| clear edge declared in the header
        ePhase := E_DL_TobCutPhase.IDLE;
    END_IF
END_IF
END_FUNCTION_BLOCK

(* ---- FB_DL_TrackBarcodeTrace.st ---- *)
//==============================================================================
// 功能块：FB_DL_TrackBarcodeTrace ｜ 中文名称：托盘条码路由追溯
// 所属子库：DL_Process ｜ 版本：v1.0.0 ｜ 兼容：CODESYS V3.5+ / TwinCAT 3 / 汇川 InoProShop
// 功能描述：托盘条码扫码路由——触发沿进扫码态，扫码枪以「bScanDone +
//           sBarcode」契约回读（R49 字符串纪律：超限截断判定在钳长
//           之前）；判据：前缀 A 匹配 → A 道、前缀 B 匹配 → B 道、
//           空码或双前缀均不匹配 → 拒收道；扫码超时（触发后超时窗满
//           bScanDone 未到）→ 故障。追溯码（sTraceCode）随路由结果
//           锁存输出，供上位追溯链消费。触发到判定的握手为单次有效
//           （bScanDone 需在触发后、超时窗内到，迟到作废）。
// 开源溯源 (Origin)：道莅原创实现（参考产线追溯与分道路由工程惯例 分类与参数域）
// 单位表：时间[ms] / 字符串长度[字符] / 道别[—]
// 错误码表：16#0005_01F6 信息级（路由判定完成：分道结果当拍有效，不置
//           bError）/ 16#0005_01F7 信息级（空码或无匹配按拒收路由降级
//           提示，不置 bError）/ 16#0005_0336 故障级（扫码超时：超时窗
//           满 bScanDone 未到，锁存，置 bError——该场景不可由 0337 的
//           组态类判据观测，属扫码枪握手独立域）/ 16#0005_0337 故障级
//           （组态非法：两前缀均为空字符串，判据无定义，置 bError）/
//           16#0005_0338 故障级兜底（状态机落 ELSE，置 bError）
// 状态机：E_DL_BarcodeRouteState（四态：eIdle=0 / eScanning=10 /
//           eRouted=20 / eFault=99），CASE 含 ELSE 兜底，ELSE 置 0338
//           并清路由输出
// 边界行为：① 组态非法（双前缀均空）→ 故障态锁存，bReset 复位；②
//           扫码态新触发沿不重置（单次握手，防连击）；③ 空码/无匹配
//           → 拒收道 + 信息 01F7 降级可观测；④ 迟到的 bScanDone（超时
//           后）作废不判（防陈旧数据误路由）；⑤ 未触发/故障态路由输出
//           清零并 bValid := FALSE；⑥ eRouted 等触发撤销回空闲（同拍
//           重启防抖，R39 范式）。
// 修订历史：v1.0.0 2026-11-17 首版（R24 派单 · ROADMAP P0 §469）
//==============================================================================

(*------------------------------------------------------------------------------
 * 枚举: E_DL_BarcodeRouteState（归属本功能块，同文件发布，全库唯一定义）
 * 含义: 扫码路由相位，每个成员在 CASE 中有且仅有一个标签。
 *-----------------------------------------------------------------------------*)
TYPE E_DL_BarcodeRouteState :
(
    eIdle     := 0,   // 空闲：等触发沿 / Idle, awaiting trigger edge
    eScanning := 10,  // 扫码：等握手或超时 / Scanning, awaiting handshake or timeout
    eRouted   := 20,  // 已路由：结果锁存，等触发撤销 / Routed, result latched, awaiting trigger drop
    eFault    := 99   // 故障：超时/组态/非法状态 / Fault, timeout, config or illegal state
);
END_TYPE

(*------------------------------------------------------------------------------
 * 枚举: E_DL_LaneRoute（归属本功能块，同文件发布，全库唯一定义）
 * 含义: 分道判定结果。
 *-----------------------------------------------------------------------------*)
TYPE E_DL_LaneRoute :
(
    eNone    := 0,   // 无判定：未路由 / None, not routed
    eLaneA   := 1,   // A 道：前缀 A 匹配 / Lane A, prefix A matched
    eLaneB   := 2,   // B 道：前缀 B 匹配 / Lane B, prefix B matched
    eReject  := 3    // 拒收道：空码或无匹配 / Reject lane, empty or unmatched
);
END_TYPE

FUNCTION_BLOCK FB_DL_TrackBarcodeTrace
VAR_INPUT
    bTrigger      : BOOL;                   // 触发扫码 [—]，上升沿生效 / Trigger scan, rising edge
    bReset        : BOOL;                   // 故障复位 [—]，上升沿清故障态 / Fault reset, rising edge clears the fault state
    sBarcode      : STRING(32);             // 扫码枪回读码 [字符]，超 32 字符截断（截断判定先于钳长，R49） / Scanner barcode [chars], truncated beyond 32
    bScanDone     : BOOL;                   // 扫码完成握手 [—]（单次有效） / Scan-done handshake, single-shot
    sRoutePrefixA : STRING(8) := 'A';       // A 道前缀 [字符]，两前缀不得均空 / Lane A prefix [chars]
    sRoutePrefixB : STRING(8) := 'B';       // B 道前缀 [字符] / Lane B prefix [chars]
    tScanTimeout  : TIME  := T#2S;          // 扫码超时窗 [ms]，须 > 0 / Scan timeout window [ms]
END_VAR
VAR_OUTPUT
    eRoute     : E_DL_LaneRoute;            // 分道判定 [—] / Lane verdict
    bLaneA     : BOOL;                      // A 道输出 [—] / Lane A output
    bLaneB     : BOOL;                      // B 道输出 [—] / Lane B output
    bReject    : BOOL;                      // 拒收道输出 [—] / Reject lane output
    sTraceCode : STRING(32);                // 追溯码 [字符]（路由结果锁存随行） / Trace code [chars], latched with the verdict
    eState     : E_DL_BarcodeRouteState;    // 相位出口 [—] / Phase outlet
    eErr       : UDINT;                     // 错误码，0 = 无错，码位 16#0005_01F6 起信息级、16#0005_0336 起故障级（分带见错误码表） / Error code, 0 = no error, band info/fault per the code table
    bError     : BOOL;                      // 故障级标志，仅故障级错误置位 / Fault-class flag, set only on fault-level codes
    bValid     : BOOL;                      // 输出可用标志 / Outputs usable flag
END_VAR
VAR
    fbTimeout : TON;                        // 扫码超时计时（每拍无条件刷新）[ms] / Scan timeout timer, refreshed unconditionally
    fbTrig    : R_TRIG;                     // 触发沿检测（待机/故障分支同样无条件刷新） / Trigger edge detector, refreshed unconditionally
    _eState   : E_DL_BarcodeRouteState := E_DL_BarcodeRouteState.eIdle; // 当前相位 / Current phase
    _bCfgBad  : BOOL;                       // 组态非法锁存 / Illegal config latch
    _eVerdict : E_DL_LaneRoute := E_DL_LaneRoute.eNone; // 判定暂存 / Verdict staging
    _sCapture : STRING(32);                 // 捕获码暂存 [字符] / Captured barcode staging [chars]
    _bInfoRoute: BOOL;                      // 判定完成信息当拍标志 / Verdict info flag of this scan
    _bInfoRej : BOOL;                       // 拒收降级信息当拍标志 / Reject-degrade info flag of this scan
    _bIllegal : BOOL;                       // 非法状态标志 / Illegal state flag
    _bInit    : BOOL := FALSE;              // 首扫标志，初值 FALSE 取非判定 / First-scan flag, tested negated
    _nLen     : INT;                        // 回读码长度 [字符] / Barcode length [chars]
END_VAR
VAR CONSTANT
    DL_TBT_STR_MAX : INT := 32;             // 追溯码容量上限 [字符] / Trace-code capacity [chars]
    DL_TBT_ZERO    : INT := 0;              // 零值常量，避免裸字面量 [字符] / Zero constant, avoids a bare literal [chars]
END_VAR

(*------------------------------------------------------------------------------
 * 段 1｜每拍预置：路由输出先清（安全侧），单拍标志预清零
 *      Route outputs cleared fail-safe first, one-shot flags pre-cleared
 *-----------------------------------------------------------------------------*)
eRoute   := E_DL_LaneRoute.eNone;        // 分道判定先清 / Verdict cleared first
bLaneA   := FALSE;                       // A 道先清 / Lane A cleared first
bLaneB   := FALSE;                       // B 道先清 / Lane B cleared first
bReject  := FALSE;                       // 拒收道先清 / Reject cleared first
sTraceCode := '';                        // 追溯码先清（路由态在段 5 重置） / Trace code cleared first
eErr   := 16#0000_0000;                  // 错误码每拍重算 / Error code recomputed
bError := FALSE;                         // 故障标志每拍重算 / Fault flag recomputed
bValid := FALSE;                         // 可用标志每拍重算 / Usable flag recomputed
_bInfoRoute := FALSE;                    // 判定信息预清零 / Verdict info pre-cleared
_bInfoRej   := FALSE;                    // 拒收信息预清零 / Reject info pre-cleared
_bIllegal   := FALSE;                    // 非法状态预清零 / Illegal flag pre-cleared

(*------------------------------------------------------------------------------
 * 段 2｜首扫初始化
 *      First-scan initialisation
 *-----------------------------------------------------------------------------*)
IF NOT _bInit THEN
    _eState  := E_DL_BarcodeRouteState.eIdle; // 相位空闲起步 / Phase starts idle
    _bCfgBad := FALSE;                   // 组态锁存清零 / Config latch cleared
    _bInit   := TRUE;                    // 首扫只做一次 / The first scan runs once
END_IF

(*------------------------------------------------------------------------------
 * 段 3｜组态闸 + 沿/超时无条件刷新（R40：CASE 之外每拍必调）
 *      Config gate plus unconditional refresh per R40
 *-----------------------------------------------------------------------------*)
fbTrig(CLK := bTrigger);                 // 触发沿检测 / Trigger edge detection
fbTimeout(IN := (_eState = E_DL_BarcodeRouteState.eScanning), PT := tScanTimeout); // 扫码超时窗 / Scan timeout window
IF (LEN(sRoutePrefixA) = DL_TBT_ZERO) AND (LEN(sRoutePrefixB) = DL_TBT_ZERO) THEN
    _bCfgBad := TRUE;                    // 双前缀均空：判据无定义锁存（0337） / Both prefixes empty, criteria undefined
END_IF
IF bReset THEN
    _bCfgBad := FALSE;                   // 复位清组态锁存 / Reset clears the config latch
END_IF

(*------------------------------------------------------------------------------
 * 段 4｜相位机（CASE 含 ELSE 兜底；状态改写只出现在分支判据内，R39）
 *      Phase machine with ELSE fallback
 *-----------------------------------------------------------------------------*)
CASE _eState OF

    E_DL_BarcodeRouteState.eIdle:          // 空闲：触发沿且组态合法进扫码
        IF fbTrig.Q AND (NOT _bCfgBad) THEN
            _eState := E_DL_BarcodeRouteState.eScanning; // 进扫码 / To scanning
        ELSIF fbTrig.Q AND _bCfgBad THEN
            _eState := E_DL_BarcodeRouteState.eFault; // 组态非法进故障 / Illegal config to fault
        END_IF

    E_DL_BarcodeRouteState.eScanning:      // 扫码：握手判定或超时
        IF _bCfgBad THEN
            _eState := E_DL_BarcodeRouteState.eFault; // 组态漂移转故障 / Config drift, fault
        ELSIF fbTimeout.Q THEN
            _eState := E_DL_BarcodeRouteState.eFault; // 超时进故障（迟到的握手作废） / Timeout to fault, late handshake void
        ELSIF bScanDone THEN
            _nLen := LEN(sBarcode);        // 回读码长度 [字符] / Barcode length
            IF _nLen = DL_TBT_ZERO THEN
                _eVerdict := E_DL_LaneRoute.eReject; // 空码拒收（R49：判定在钳长前） / Empty barcode, reject
                _bInfoRej := TRUE;         // 拒收降级提示（信息级） / Reject-degrade notice, info
            ELSE
                IF _nLen > DL_TBT_STR_MAX THEN
                    _nLen := DL_TBT_STR_MAX; // 超限先置截断判定再钳长（本件容量即 32，防御路径） / Truncation verdict before the clamp per R49
                    _bInfoRej := TRUE;     // 截断归拒收降级提示（信息级） / Truncation folded into the degrade notice
                END_IF
                _sCapture := LEFT(sBarcode, _nLen); // 钳长后捕获 / Captured after the clamp
                IF (LEN(sRoutePrefixA) > DL_TBT_ZERO)
                   AND (LEFT(_sCapture, LEN(sRoutePrefixA)) = sRoutePrefixA) THEN
                    _eVerdict := E_DL_LaneRoute.eLaneA; // 前缀 A 匹配 → A 道 / Prefix A matched
                ELSIF (LEN(sRoutePrefixB) > DL_TBT_ZERO)
                   AND (LEFT(_sCapture, LEN(sRoutePrefixB)) = sRoutePrefixB) THEN
                    _eVerdict := E_DL_LaneRoute.eLaneB; // 前缀 B 匹配 → B 道 / Prefix B matched
                ELSE
                    _eVerdict := E_DL_LaneRoute.eReject; // 无匹配拒收 / No match, reject
                    _bInfoRej := TRUE;     // 拒收降级提示（信息级） / Reject-degrade notice, info
                END_IF
            END_IF
            _eState := E_DL_BarcodeRouteState.eRouted; // 进路由态锁存 / To routed, latched
        END_IF

    E_DL_BarcodeRouteState.eRouted:        // 已路由：等触发撤销回空闲（同拍重启防抖）
        IF NOT bTrigger THEN
            _eVerdict := E_DL_LaneRoute.eNone; // 判定复位 / Verdict reset
            _eState := E_DL_BarcodeRouteState.eIdle; // 回空闲 / Back to idle
        END_IF

    E_DL_BarcodeRouteState.eFault:         // 故障：复位沿且原因消失回空闲
        IF bReset AND (NOT _bCfgBad) THEN
            _eState := E_DL_BarcodeRouteState.eIdle; // 回空闲 / Back to idle
        END_IF

    ELSE                                   // 非法状态兜底（R21：CASE 必带 ELSE）
        _bIllegal := TRUE;                 // 标记非法状态 / Flag the illegal state
        _eVerdict := E_DL_LaneRoute.eNone; // 判定复位 / Verdict reset
        _eState := E_DL_BarcodeRouteState.eFault; // 回故障态 / Back to fault
END_CASE

(*------------------------------------------------------------------------------
 * 段 5｜路由出口（eRouted 态单源赋值；互斥由 IF/ELSE 结构性成立）
 *      Route outlet, single-source in the routed phase
 *-----------------------------------------------------------------------------*)
CASE _eVerdict OF
    E_DL_LaneRoute.eLaneA:                 // A 道 / Lane A
        bLaneA := TRUE;                    // A 道输出 / Lane A output
    E_DL_LaneRoute.eLaneB:                 // B 道 / Lane B
        bLaneB := TRUE;                    // B 道输出 / Lane B output
    E_DL_LaneRoute.eReject:                // 拒收道 / Reject lane
        bReject := TRUE;                   // 拒收道输出 / Reject output
    ELSE                                   // 无判定：输出全清 / No verdict, all clear
        _eVerdict := _eVerdict;            // 保持预置清零（判定维持空档，显式自持）/ Stays cleared (explicit self-hold)
END_CASE
IF _eState = E_DL_BarcodeRouteState.eRouted THEN
    eRoute := _eVerdict;                   // 判定出口（路由态） / Verdict outlet in the routed phase
    IF _eVerdict <> E_DL_LaneRoute.eNone THEN
        sTraceCode := _sCapture;           // 追溯码随行（仅有效判定） / Trace code attached to a valid verdict
        _bInfoRoute := TRUE;               // 判定完成信息（信息级） / Verdict-done info
    END_IF
END_IF

(*------------------------------------------------------------------------------
 * 段 6｜码位出口与放行（故障级码 3 行内置 bError，R45/R101 配对）
 *      Code outlet and release, fault codes paired with bError
 *-----------------------------------------------------------------------------*)
IF _bIllegal THEN
    eErr   := 16#0005_0338;                // 故障级：状态机兜底 / Fault: state machine fallback
    bError := TRUE;                        // 置故障标志 / Raise the fault flag
ELSIF _bCfgBad THEN
    eErr   := 16#0005_0337;                // 故障级：组态非法（双前缀均空） / Fault: illegal configuration
    bError := TRUE;                        // 置故障标志 / Raise the fault flag
ELSIF (_eState = E_DL_BarcodeRouteState.eFault) AND (NOT _bCfgBad) THEN
    eErr   := 16#0005_0336;                // 故障级：扫码超时 / Fault: scan timeout
    bError := TRUE;                        // 置故障标志 / Raise the fault flag
ELSIF _bInfoRej THEN
    eErr := 16#0005_01F7;                  // 信息级：空码/无匹配/截断按拒收降级 / Info: reject-degrade notice
ELSIF _bInfoRoute THEN
    eErr := 16#0005_01F6;                  // 信息级：路由判定完成 / Info: verdict done
END_IF

bValid := (NOT bError) AND (_eState = E_DL_BarcodeRouteState.eRouted); // 仅路由态放行 / Usable only in the routed phase
eState := _eState;                       // 相位出口 / Phase outlet
END_FUNCTION_BLOCK

(* ---- FB_DL_TrackerWindStow.st ---- *)
(*
  FB_DL_TrackerWindStow  —  跟踪支架大风保护收拢 / Tracker wind-stow protection
  分类 Category : DL_Process
  码位 Code     : 16#06_0_8C
  版本 Version  : 1.0.0
  溯源 Source   : LGF Technology 语义借鉴 · clean-room 实现，仅借分类/参数域/命名，未复制源码
  功能 Function : 1) 风速超「高阈值（带迟滞）」或趋势判据（风速爬升率超限持续 N 拍）→ 置收拢命令；
                  2) 解除条件：风速回落到解除阈值以下 + 最短驻留时间到 → 自动解除（解除路径可达）；
                  3) 收拢角度命令钳位到行程域，防组态越程。
  边界 Boundary : ① 风速非有限或 < 0 判无效：冻结输出保持末次命令并置信息码；
                  ② 高/解除阈值倒置或爬升率门限 <= 0 出厂报码不运行（组态闸）；
                  ③ 趋势窗确认拍数不足不出趋势结论（N 拍未满不参与判据）；
                  ④ 输出三行同向：收拢命令 → 安全角度 → 趋势告警标志。
  依赖 Depends  : FB_DL_Differentiator（风速爬升率，每拍无条件调用）

  码表 Error codes（本件子码步进 16#10，避让邻件码位）:
    16#0002_068C 故障级：组态非法（高/解除阈值倒置、爬升率门限 <= 0、收拢角行程域倒置）
    16#0002_069C 故障级：相 ID 越界（枚举兜底路径）
    16#0002_06AC 信息级：风速无效冻结输出 / 趋势确认拍数不足不出结论（不置 bError）
*)

TYPE E_DL_TwsPhase :
(
    eIdle    := 0,   // 空闲待机 / Idle
    eMonitor := 10,  // 风况监视 / Wind monitoring
    eStow    := 20,  // 大风收拢命令保持 / Stow command held
    eRelease := 30,  // 解除驻留等待（风速已回落）/ Release dwell after wind dropped
    eFrozen  := 40,  // 风速无效冻结 / Frozen by invalid wind
    eFault   := 90   // 组态故障锁定 / Configuration fault locked
);
END_TYPE

FUNCTION_BLOCK FB_DL_TrackerWindStow
VAR_INPUT
    bEnable        : BOOL;                          // 总使能，FALSE 回空闲 / Master enable
    bReset         : BOOL;                          // 复位，上升沿清组态故障 / Reset, clears configuration fault
    fWindSpeed     : REAL;                          // 风速实测 [m/s]，域 >= 0 / Measured wind speed [m/s]
    fWindHigh      : REAL := 25.0;                  // 大风收拢阈值 [m/s]，须 > 解除阈值 / Stow threshold [m/s]
    fWindRelease   : REAL := 18.0;                  // 解除阈值 [m/s]，带迟滞 / Release threshold [m/s]
    fRiseRateMax   : REAL := 2.0;                   // 风速爬升率门限 [m/s per s]，域 > 0 / Rise-rate limit [m/s per s]
    uRiseConfirm   : UINT := 5;                     // 趋势确认拍数 [拍]，0 = 禁用趋势判据 / Trend confirm scans [scan]
    fStowAngle     : REAL := 60.0;                  // 安全收拢角度 [deg] / Safety stow angle [deg]
    fAngleMax      : REAL := 75.0;                  // 行程域上限 [deg]，收拢角钳位域 / Travel domain high [deg]
    fAngleMin      : REAL := -75.0;                 // 行程域下限 [deg] / Travel domain low [deg]
    fDwellSec      : REAL := 30.0;                  // 解除最短驻留 [s]，域 > 0 / Min release dwell [s]
    fTaskCycle     : REAL := 0.1;                   // 任务周期 [s]，域 > 0 / Task cycle [s]
    fEps           : REAL := 1.0E-6;                // 浮点判零容差 [1] / Floating zero tolerance
END_VAR
VAR_OUTPUT
    bStowCmd       : BOOL;                          // 收拢命令出口（保持型）/ Stow command output, held
    fStowAngleCmd  : REAL;                          // 安全角度命令 [deg]，已钳行程域 / Safe angle command [deg], clamped
    bTrendAlarm    : BOOL;                          // 趋势判据命中标志（本拍重算）/ Trend criterion hit flag
    bFrozen        : BOOL;                          // 冻结标志（风速无效）/ Frozen by invalid wind
    bError         : BOOL;                          // 故障标志，与故障级码配对 / Fault flag paired with fault codes
    uErrorId       : UDINT;                         // 事件码，0 = 无事件 / Event code, 0 = none
    eStateOut      : E_DL_TwsPhase;                 // 状态机当前态，段尾单点映射 / Phase mapped at tail
END_VAR
VAR
    _eState        : E_DL_TwsPhase := E_DL_TwsPhase.eIdle;  // 内部状态 / Internal state
    fbDiff         : FB_DL_Differentiator;          // 风速爬升率实例（无条件调用）/ Rise-rate instance
    rtrReset       : R_TRIG;                        // 复位沿 / Reset edge
    rtrWindOk      : R_TRIG;                        // 风速恢复沿（解除冻结重计驻留）/ Wind-valid edge
    tonDwell       : TON;                           // 解除驻留定时器（IN := NOT Q 自复位见 R33-2 用法不适用，此处电平触发）/ Release dwell timer
    bCfgOk         : BOOL;                          // 组态合法标志 / Configuration valid
    bWindOk        : BOOL;                          // 本拍风速有效 / Wind valid this scan
    bOverHigh      : BOOL;                          // 超高阈值（电平）/ Above stow threshold, level
    bBelowRelease  : BOOL;                          // 低于解除阈值（电平）/ Below release threshold, level
    bTrendHit      : BOOL;                          // 趋势判据命中（电平）/ Trend criterion hit
    uTrendCnt      : UINT;                          // 趋势确认计数 [拍] / Trend confirm counter [scan]
    fRateEff       : REAL;                          // 本拍爬升率 [m/s per s] / Rise rate this scan [m/s per s]
    uFault         : UDINT;                         // 锁存故障码 / Latched fault code
    uInfo          : UDINT;                         // 信息级码（本拍重算）/ Information code
END_VAR
VAR CONSTANT
    DL_TWS_INF_MAX : REAL := 1.0E30;                // 有限值判定幅值上限 [m/s] / Finite magnitude bound [m/s]
    DL_TWS_ANG_MAX : REAL := 180.0;                 // 角度物理域上限 [deg] / Angle domain high [deg]
END_VAR

(* === 段 0 · 实例刷新（无条件周期调用）=== *)
rtrReset(CLK := bReset);                          // 每拍刷新复位沿
rtrWindOk(CLK := bWindOk);                        // 每拍刷新风速恢复沿
fbDiff(bEnable := bCfgOk AND bEnable,             // 组态闸过才使能微分（每拍仍无条件调用实例）
       fIn := fWindSpeed,                         // 被微分量为风速
       tFiltTime := T#2S,                         // 爬升率低通 2 s 抑制阵风毛刺
       tSampleTime := REAL_TO_TIME(MAX(fTaskCycle, 0.01) * 1000.0),  // 周期换算 [ms]
       rRateMax := 1.0E10,                        // 速率上限放开，门限由本件判
       rRateMin := -1.0E10);                      // 速率下限放开

(* === 段 1 · 组态闸与输入域闸 === *)
bCfgOk := (fWindHigh > fWindRelease + fEps)       // 高阈值须高于解除阈值（迟滞带为正）
          AND (fWindHigh > fEps) AND (fWindRelease > fEps)
          AND (fRiseRateMax > fEps) AND (fDwellSec > fEps) AND (fTaskCycle > fEps)
          AND (fAngleMax > fAngleMin + fEps)      // 行程域不倒置
          AND (fWindHigh = fWindHigh) AND (fStowAngle = fStowAngle);  // NaN 自反
IF NOT bCfgOk THEN
    uFault := 16#0002_068C;                       // 故障级：组态非法
END_IF
IF rtrReset.Q AND bCfgOk THEN
    uFault := 16#0000;                            // 复位沿清锁存（解除路径可达）
END_IF
uInfo := 16#0000;                                 // 信息码每拍清零（R189：信息级可每拍重算）
bWindOk := (fWindSpeed = fWindSpeed) AND (fWindSpeed >= 0.0)
           AND (fWindSpeed < DL_TWS_INF_MAX);     // NaN 自反 + 非负域 + 幅值闸
IF NOT bWindOk THEN
    uInfo := 16#0002_06AC;                        // 信息级：风速无效冻结
END_IF
fStowAngleCmd := fStowAngle;                      // 角度命令先取组态值
IF fStowAngleCmd > fAngleMax THEN
    fStowAngleCmd := fAngleMax;                   // 钳到行程域上限
END_IF
IF fStowAngleCmd < fAngleMin THEN
    fStowAngleCmd := fAngleMin;                   // 钳到行程域下限
END_IF
IF ABS(fStowAngleCmd) > DL_TWS_ANG_MAX THEN
    fStowAngleCmd := 0.0;                         // 钳位后仍越物理域：安全侧回 0 度
END_IF

(* === 段 2 · 风况判据（本拍重算，非锁存）=== *)
bOverHigh := bWindOk AND (fWindSpeed >= fWindHigh);             // 电平判据：超高阈值
bBelowRelease := bWindOk AND (fWindSpeed <= fWindRelease);      // 电平判据：低于解除阈值
bTrendHit := FALSE;                                             // 趋势结论默认不成立
IF bWindOk AND fbDiff.bValid THEN
    fRateEff := fbDiff.fRateOut;                  // 取滤波后爬升率
    IF (uRiseConfirm > UINT#0) AND (fRateEff >= fRiseRateMax) THEN
        uTrendCnt := uTrendCnt + UINT#1;          // 命中拍计数累加
        IF uTrendCnt >= uRiseConfirm THEN
            bTrendHit := TRUE;                    // 连续 N 拍超门限：趋势结论成立
        END_IF
    ELSE
        uTrendCnt := UINT#0;                      // 未命中：确认计数归零重计
    END_IF
ELSE
    uTrendCnt := UINT#0;                          // 风速无效/微分未就绪：不出趋势结论
    IF bCfgOk AND (uRiseConfirm > UINT#0) THEN
        uInfo := 16#0002_06AC;                    // 信息级：趋势窗确认拍数不足不出结论
    END_IF
END_IF
bTrendAlarm := bTrendHit;                         // 趋势告警出口（本拍重算）

(* === 段 3 · 主状态机（ENUM + CASE，含 ELSE 兜底）=== *)
tonDwell(IN := (_eState = E_DL_TwsPhase.eRelease) AND bBelowRelease,   // 驻留计时只在解除相且风已回落
         PT := REAL_TO_TIME(fDwellSec * 1000.0));                      // 驻留时长换算 [ms]
CASE _eState OF
E_DL_TwsPhase.eIdle :
    bStowCmd := FALSE;                            // 空闲不收拢
    IF uFault <> 16#0000 THEN
        _eState := E_DL_TwsPhase.eFault;          // 故障优先
    ELSIF NOT bEnable THEN
        _eState := E_DL_TwsPhase.eIdle;           // 失能保持空闲
    ELSIF NOT bWindOk THEN
        _eState := E_DL_TwsPhase.eFrozen;         // 风速无效进冻结
    ELSIF bOverHigh OR bTrendHit THEN
        _eState := E_DL_TwsPhase.eStow;           // 阈值或趋势任一命中：收拢
    ELSE
        _eState := E_DL_TwsPhase.eMonitor;        // 正常进入监视相
    END_IF

E_DL_TwsPhase.eMonitor :
    bStowCmd := FALSE;                            // 监视相不收拢
    IF (NOT bWindOk) OR (uFault <> 16#0000) THEN
        _eState := E_DL_TwsPhase.eFrozen;         // 无效/故障转冻结
    ELSIF bOverHigh OR bTrendHit THEN
        _eState := E_DL_TwsPhase.eStow;           // 命中转收拢
    END_IF

E_DL_TwsPhase.eStow :
    bStowCmd := TRUE;                             // 收拢命令保持（同拍抹除防护：仅解除相清）
    IF NOT bWindOk THEN
        _eState := E_DL_TwsPhase.eFrozen;         // 收拢中风速无效：冻结保持命令
    ELSIF bBelowRelease THEN
        _eState := E_DL_TwsPhase.eRelease;        // 风已回落：进解除驻留相
    END_IF

E_DL_TwsPhase.eRelease :
    bStowCmd := TRUE;                             // 驻留期内命令仍保持（防回弹抖动）
    IF NOT bWindOk THEN
        _eState := E_DL_TwsPhase.eFrozen;         // 驻留中风速无效：冻结保持命令
    ELSIF bOverHigh OR bTrendHit THEN
        _eState := E_DL_TwsPhase.eStow;           // 风复起：回到收拢相（驻留定时器由 IN 条件自清）
    ELSIF tonDwell.Q THEN
        bStowCmd := FALSE;                        // 驻留满且风持续回落：解除命令
        uTrendCnt := UINT#0;                      // 趋势计数同步清零
        _eState := E_DL_TwsPhase.eMonitor;        // 回监视相（解除路径可达）
    END_IF

E_DL_TwsPhase.eFrozen :
    bFrozen := TRUE;                              // 冻结标志保持
    (* 收拢命令为输出保持量：冻结期间不清零，恢复后按状态续判 *)
    IF bWindOk AND (uFault = 16#0000) THEN
        bFrozen := FALSE;                         // 风速恢复：解冻（可到达的解除路径）
        IF rtrWindOk.Q THEN
            uTrendCnt := UINT#0;                  // 恢复沿重计趋势确认
        END_IF
        _eState := E_DL_TwsPhase.eMonitor;        // 回监视相
    END_IF

E_DL_TwsPhase.eFault :
    bFrozen := TRUE;                              // 故障态冻结
    bStowCmd := TRUE;                             // 故障安全侧：保持收拢命令
    IF uFault = 16#0000 THEN
        _eState := E_DL_TwsPhase.eIdle;           // 解锁回空闲
    END_IF

ELSE
    _eState := E_DL_TwsPhase.eFault;              // 非法状态拦截
    uFault := 16#0002_069C;                       // 故障级：相 ID 越界
    bFrozen := TRUE;                              // 安全侧冻结
    bStowCmd := TRUE;                             // 安全侧保持收拢
END_CASE

(* === 段 4 · 输出映射 === *)
bFrozen := (_eState = E_DL_TwsPhase.eFrozen) OR (_eState = E_DL_TwsPhase.eFault);  // 冻结标志段尾单点映射
bError := (uFault <> 16#0000);                    // 故障标志仅由故障级码置位（R45 配对）
IF bError THEN
    uErrorId := uFault;                           // 故障级优先上报
ELSE
    uErrorId := uInfo;                            // 否则上报信息级码
END_IF
eStateOut := _eState;                             // 输出枚举段尾单点映射（N2 规则）
END_FUNCTION_BLOCK
